   AryTypePara[234].Other.FixtureEnable := FALSE;
   AryTypePara[234].Other.Byte_1 := 16#00;
   AryTypePara[234].Other.Int_1 := 0;
   AryTypePara[234].Other."Char" := ' ';
   AryTypePara[234].Other.Word_1 := 16#0000;
   AryTypePara[234].Other.DInt_1 := 0;
   AryTypePara[234].Other.DWord_1 := 16#0000_0000;
   AryTypePara[234].Other.Real_1 := 0.0;
   AryTypePara[234].Other.S5Time := T#0MS;
   AryTypePara[234].Other."String" := '';
   AryTypePara[235].TypeName := '';
   AryTypePara[235].bit.Bit0 := FALSE;
   AryTypePara[235].bit.sp := 16#0000;
   AryTypePara[235].bit.Other.Bool_1 := FALSE;
   AryTypePara[235].bit.Other.Byte_2 := 16#00;
   AryTypePara[235].bit.Other.Int_1 := 0;
   AryTypePara[235].bit.Other."Char" := ' ';
   AryTypePara[235].Other.STxxxCCDProgNO := 0;
   AryTypePara[235].Other.FixtureEnable := FALSE;
   AryTypePara[235].Other.Byte_1 := 16#00;
   AryTypePara[235].Other.Int_1 := 0;
   AryTypePara[235].Other."Char" := ' ';
   AryTypePara[235].Other.Word_1 := 16#0000;
   AryTypePara[235].Other.DInt_1 := 0;
   AryTypePara[235].Other.DWord_1 := 16#0000_0000;
   AryTypePara[235].Other.Real_1 := 0.0;
   AryTypePara[235].Other.S5Time := T#0MS;
   AryTypePara[235].Other."String" := '';
   AryTypePara[236].TypeName := '';
   AryTypePara[236].bit.Bit0 := FALSE;
   AryTypePara[236].bit.sp := 16#0000;
   AryTypePara[236].bit.Other.Bool_1 := FALSE;
   AryTypePara[236].bit.Other.Byte_2 := 16#00;
   AryTypePara[236].bit.Other.Int_1 := 0;
   AryTypePara[236].bit.Other."Char" := ' ';
   AryTypePara[236].Other.STxxxCCDProgNO := 0;
   AryTypePara[236].Other.FixtureEnable := FALSE;
   AryTypePara[236].Other.Byte_1 := 16#00;
   AryTypePara[236].Other.Int_1 := 0;
   AryTypePara[236].Other."Char" := ' ';
   AryTypePara[236].Other.Word_1 := 16#0000;
   AryTypePara[236].Other.DInt_1 := 0;
   AryTypePara[236].Other.DWord_1 := 16#0000_0000;
   AryTypePara[236].Other.Real_1 := 0.0;
   AryTypePara[236].Other.S5Time := T#0MS;
   AryTypePara[236].Other."String" := '';
   AryTypePara[237].TypeName := '';
   AryTypePara[237].bit.Bit0 := FALSE;
   AryTypePara[237].bit.sp := 16#0000;
   AryTypePara[237].bit.Other.Bool_1 := FALSE;
   AryTypePara[237].bit.Other.Byte_2 := 16#00;
   AryTypePara[237].bit.Other.Int_1 := 0;
   AryTypePara[237].bit.Other."Char" := ' ';
   AryTypePara[237].Other.STxxxCCDProgNO := 0;
   AryTypePara[237].Other.FixtureEnable := FALSE;
   AryTypePara[237].Other.Byte_1 := 16#00;
   AryTypePara[237].Other.Int_1 := 0;
   AryTypePara[237].Other."Char" := ' ';
   AryTypePara[237].Other.Word_1 := 16#0000;
   AryTypePara[237].Other.DInt_1 := 0;
   AryTypePara[237].Other.DWord_1 := 16#0000_0000;
   AryTypePara[237].Other.Real_1 := 0.0;
   AryTypePara[237].Other.S5Time := T#0MS;
   AryTypePara[237].Other."String" := '';
   AryTypePara[238].TypeName := '';
   AryTypePara[238].bit.Bit0 := FALSE;
   AryTypePara[238].bit.sp := 16#0000;
   AryTypePara[238].bit.Other.Bool_1 := FALSE;
   AryTypePara[238].bit.Other.Byte_2 := 16#00;
   AryTypePara[238].bit.Other.Int_1 := 0;
   AryTypePara[238].bit.Other."Char" := ' ';
   AryTypePara[238].Other.STxxxCCDProgNO := 0;
   AryTypePara[238].Other.FixtureEnable := FALSE;
   AryTypePara[238].Other.Byte_1 := 16#00;
   AryTypePara[238].Other.Int_1 := 0;
   AryTypePara[238].Other."Char" := ' ';
   AryTypePara[238].Other.Word_1 := 16#0000;
   AryTypePara[238].Other.DInt_1 := 0;
   AryTypePara[238].Other.DWord_1 := 16#0000_0000;
   AryTypePara[238].Other.Real_1 := 0.0;
   AryTypePara[238].Other.S5Time := T#0MS;
   AryTypePara[238].Other."String" := '';
   AryTypePara[239].TypeName := '';
   AryTypePara[239].bit.Bit0 := FALSE;
   AryTypePara[239].bit.sp := 16#0000;
   AryTypePara[239].bit.Other.Bool_1 := FALSE;
   AryTypePara[239].bit.Other.Byte_2 := 16#00;
   AryTypePara[239].bit.Other.Int_1 := 0;
   AryTypePara[239].bit.Other."Char" := ' ';
   AryTypePara[239].Other.STxxxCCDProgNO := 0;
   AryTypePara[239].Other.FixtureEnable := FALSE;
   AryTypePara[239].Other.Byte_1 := 16#00;
   AryTypePara[239].Other.Int_1 := 0;
   AryTypePara[239].Other."Char" := ' ';
   AryTypePara[239].Other.Word_1 := 16#0000;
   AryTypePara[239].Other.DInt_1 := 0;
   AryTypePara[239].Other.DWord_1 := 16#0000_0000;
   AryTypePara[239].Other.Real_1 := 0.0;
   AryTypePara[239].Other.S5Time := T#0MS;
   AryTypePara[239].Other."String" := '';
   AryTypePara[240].TypeName := '';
   AryTypePara[240].bit.Bit0 := FALSE;
   AryTypePara[240].bit.sp := 16#0000;
   AryTypePara[240].bit.Other.Bool_1 := FALSE;
   AryTypePara[240].bit.Other.Byte_2 := 16#00;
   AryTypePara[240].bit.Other.Int_1 := 0;
   AryTypePara[240].bit.Other."Char" := ' ';
   AryTypePara[240].Other.STxxxCCDProgNO := 0;
   AryTypePara[240].Other.FixtureEnable := FALSE;
   AryTypePara[240].Other.Byte_1 := 16#00;
   AryTypePara[240].Other.Int_1 := 0;
   AryTypePara[240].Other."Char" := ' ';
   AryTypePara[240].Other.Word_1 := 16#0000;
   AryTypePara[240].Other.DInt_1 := 0;
   AryTypePara[240].Other.DWord_1 := 16#0000_0000;
   AryTypePara[240].Other.Real_1 := 0.0;
   AryTypePara[240].Other.S5Time := T#0MS;
   AryTypePara[240].Other."String" := '';
   AryTypePara[241].TypeName := '';
   AryTypePara[241].bit.Bit0 := FALSE;
   AryTypePara[241].bit.sp := 16#0000;
   AryTypePara[241].bit.Other.Bool_1 := FALSE;
   AryTypePara[241].bit.Other.Byte_2 := 16#00;
   AryTypePara[241].bit.Other.Int_1 := 0;
   AryTypePara[241].bit.Other."Char" := ' ';
   AryTypePara[241].Other.STxxxCCDProgNO := 0;
   AryTypePara[241].Other.FixtureEnable := FALSE;
   AryTypePara[241].Other.Byte_1 := 16#00;
   AryTypePara[241].Other.Int_1 := 0;
   AryTypePara[241].Other."Char" := ' ';
   AryTypePara[241].Other.Word_1 := 16#0000;
   AryTypePara[241].Other.DInt_1 := 0;
   AryTypePara[241].Other.DWord_1 := 16#0000_0000;
   AryTypePara[241].Other.Real_1 := 0.0;
   AryTypePara[241].Other.S5Time := T#0MS;
   AryTypePara[241].Other."String" := '';
   AryTypePara[242].TypeName := '';
   AryTypePara[242].bit.Bit0 := FALSE;
   AryTypePara[242].bit.sp := 16#0000;
   AryTypePara[242].bit.Other.Bool_1 := FALSE;
   AryTypePara[242].bit.Other.Byte_2 := 16#00;
   AryTypePara[242].bit.Other.Int_1 := 0;
   AryTypePara[242].bit.Other."Char" := ' ';
   AryTypePara[242].Other.STxxxCCDProgNO := 0;
   AryTypePara[242].Other.FixtureEnable := FALSE;
   AryTypePara[242].Other.Byte_1 := 16#00;
   AryTypePara[242].Other.Int_1 := 0;
   AryTypePara[242].Other."Char" := ' ';
   AryTypePara[242].Other.Word_1 := 16#0000;
   AryTypePara[242].Other.DInt_1 := 0;
   AryTypePara[242].Other.DWord_1 := 16#0000_0000;
   AryTypePara[242].Other.Real_1 := 0.0;
   AryTypePara[242].Other.S5Time := T#0MS;
   AryTypePara[242].Other."String" := '';
   AryTypePara[243].TypeName := '';
   AryTypePara[243].bit.Bit0 := FALSE;
   AryTypePara[243].bit.sp := 16#0000;
   AryTypePara[243].bit.Other.Bool_1 := FALSE;
   AryTypePara[243].bit.Other.Byte_2 := 16#00;
   AryTypePara[243].bit.Other.Int_1 := 0;
   AryTypePara[243].bit.Other."Char" := ' ';
   AryTypePara[243].Other.STxxxCCDProgNO := 0;
   AryTypePara[243].Other.FixtureEnable := FALSE;
   AryTypePara[243].Other.Byte_1 := 16#00;
   AryTypePara[243].Other.Int_1 := 0;
   AryTypePara[243].Other."Char" := ' ';
   AryTypePara[243].Other.Word_1 := 16#0000;
   AryTypePara[243].Other.DInt_1 := 0;
   AryTypePara[243].Other.DWord_1 := 16#0000_0000;
   AryTypePara[243].Other.Real_1 := 0.0;
   AryTypePara[243].Other.S5Time := T#0MS;
   AryTypePara[243].Other."String" := '';
   AryTypePara[244].TypeName := '';
   AryTypePara[244].bit.Bit0 := FALSE;
   AryTypePara[244].bit.sp := 16#0000;
   AryTypePara[244].bit.Other.Bool_1 := FALSE;
   AryTypePara[244].bit.Other.Byte_2 := 16#00;
   AryTypePara[244].bit.Other.Int_1 := 0;
   AryTypePara[244].bit.Other."Char" := ' ';
   AryTypePara[244].Other.STxxxCCDProgNO := 0;
   AryTypePara[244].Other.FixtureEnable := FALSE;
   AryTypePara[244].Other.Byte_1 := 16#00;
   AryTypePara[244].Other.Int_1 := 0;
   AryTypePara[244].Other."Char" := ' ';
   AryTypePara[244].Other.Word_1 := 16#0000;
   AryTypePara[244].Other.DInt_1 := 0;
   AryTypePara[244].Other.DWord_1 := 16#0000_0000;
   AryTypePara[244].Other.Real_1 := 0.0;
   AryTypePara[244].Other.S5Time := T#0MS;
   AryTypePara[244].Other."String" := '';
   AryTypePara[245].TypeName := '';
   AryTypePara[245].bit.Bit0 := FALSE;
   AryTypePara[245].bit.sp := 16#0000;
   AryTypePara[245].bit.Other.Bool_1 := FALSE;
   AryTypePara[245].bit.Other.Byte_2 := 16#00;
   AryTypePara[245].bit.Other.Int_1 := 0;
   AryTypePara[245].bit.Other."Char" := ' ';
   AryTypePara[245].Other.STxxxCCDProgNO := 0;
   AryTypePara[245].Other.FixtureEnable := FALSE;
   AryTypePara[245].Other.Byte_1 := 16#00;
   AryTypePara[245].Other.Int_1 := 0;
   AryTypePara[245].Other."Char" := ' ';
   AryTypePara[245].Other.Word_1 := 16#0000;
   AryTypePara[245].Other.DInt_1 := 0;
   AryTypePara[245].Other.DWord_1 := 16#0000_0000;
   AryTypePara[245].Other.Real_1 := 0.0;
   AryTypePara[245].Other.S5Time := T#0MS;
   AryTypePara[245].Other."String" := '';
   AryTypePara[246].TypeName := '';
   AryTypePara[246].bit.Bit0 := FALSE;
   AryTypePara[246].bit.sp := 16#0000;
   AryTypePara[246].bit.Other.Bool_1 := FALSE;
   AryTypePara[246].bit.Other.Byte_2 := 16#00;
   AryTypePara[246].bit.Other.Int_1 := 0;
   AryTypePara[246].bit.Other."Char" := ' ';
   AryTypePara[246].Other.STxxxCCDProgNO := 0;
   AryTypePara[246].Other.FixtureEnable := FALSE;
   AryTypePara[246].Other.Byte_1 := 16#00;
   AryTypePara[246].Other.Int_1 := 0;
   AryTypePara[246].Other."Char" := ' ';
   AryTypePara[246].Other.Word_1 := 16#0000;
   AryTypePara[246].Other.DInt_1 := 0;
   AryTypePara[246].Other.DWord_1 := 16#0000_0000;
   AryTypePara[246].Other.Real_1 := 0.0;
   AryTypePara[246].Other.S5Time := T#0MS;
   AryTypePara[246].Other."String" := '';
   AryTypePara[247].TypeName := '';
   AryTypePara[247].bit.Bit0 := FALSE;
   AryTypePara[247].bit.sp := 16#0000;
   AryTypePara[247].bit.Other.Bool_1 := FALSE;
   AryTypePara[247].bit.Other.Byte_2 := 16#00;
   AryTypePara[247].bit.Other.Int_1 := 0;
   AryTypePara[247].bit.Other."Char" := ' ';
   AryTypePara[247].Other.STxxxCCDProgNO := 0;
   AryTypePara[247].Other.FixtureEnable := FALSE;
   AryTypePara[247].Other.Byte_1 := 16#00;
   AryTypePara[247].Other.Int_1 := 0;
   AryTypePara[247].Other."Char" := ' ';
   AryTypePara[247].Other.Word_1 := 16#0000;
   AryTypePara[247].Other.DInt_1 := 0;
   AryTypePara[247].Other.DWord_1 := 16#0000_0000;
   AryTypePara[247].Other.Real_1 := 0.0;
   AryTypePara[247].Other.S5Time := T#0MS;
   AryTypePara[247].Other."String" := '';
   AryTypePara[248].TypeName := '';
   AryTypePara[248].bit.Bit0 := FALSE;
   AryTypePara[248].bit.sp := 16#0000;
   AryTypePara[248].bit.Other.Bool_1 := FALSE;
   AryTypePara[248].bit.Other.Byte_2 := 16#00;
   AryTypePara[248].bit.Other.Int_1 := 0;
   AryTypePara[248].bit.Other."Char" := ' ';
   AryTypePara[248].Other.STxxxCCDProgNO := 0;
   AryTypePara[248].Other.FixtureEnable := FALSE;
   AryTypePara[248].Other.Byte_1 := 16#00;
   AryTypePara[248].Other.Int_1 := 0;
   AryTypePara[248].Other."Char" := ' ';
   AryTypePara[248].Other.Word_1 := 16#0000;
   AryTypePara[248].Other.DInt_1 := 0;
   AryTypePara[248].Other.DWord_1 := 16#0000_0000;
   AryTypePara[248].Other.Real_1 := 0.0;
   AryTypePara[248].Other.S5Time := T#0MS;
   AryTypePara[248].Other."String" := '';
   AryTypePara[249].TypeName := '';
   AryTypePara[249].bit.Bit0 := FALSE;
   AryTypePara[249].bit.sp := 16#0000;
   AryTypePara[249].bit.Other.Bool_1 := FALSE;
   AryTypePara[249].bit.Other.Byte_2 := 16#00;
   AryTypePara[249].bit.Other.Int_1 := 0;
   AryTypePara[249].bit.Other."Char" := ' ';
   AryTypePara[249].Other.STxxxCCDProgNO := 0;
   AryTypePara[249].Other.FixtureEnable := FALSE;
   AryTypePara[249].Other.Byte_1 := 16#00;
   AryTypePara[249].Other.Int_1 := 0;
   AryTypePara[249].Other."Char" := ' ';
   AryTypePara[249].Other.Word_1 := 16#0000;
   AryTypePara[249].Other.DInt_1 := 0;
   AryTypePara[249].Other.DWord_1 := 16#0000_0000;
   AryTypePara[249].Other.Real_1 := 0.0;
   AryTypePara[249].Other.S5Time := T#0MS;
   AryTypePara[249].Other."String" := '';
   AryTypePara[250].TypeName := '';
   AryTypePara[250].bit.Bit0 := FALSE;
   AryTypePara[250].bit.sp := 16#0000;
   AryTypePara[250].bit.Other.Bool_1 := FALSE;
   AryTypePara[250].bit.Other.Byte_2 := 16#00;
   AryTypePara[250].bit.Other.Int_1 := 0;
   AryTypePara[250].bit.Other."Char" := ' ';
   AryTypePara[250].Other.STxxxCCDProgNO := 0;
   AryTypePara[250].Other.FixtureEnable := FALSE;
   AryTypePara[250].Other.Byte_1 := 16#00;
   AryTypePara[250].Other.Int_1 := 0;
   AryTypePara[250].Other."Char" := ' ';
   AryTypePara[250].Other.Word_1 := 16#0000;
   AryTypePara[250].Other.DInt_1 := 0;
   AryTypePara[250].Other.DWord_1 := 16#0000_0000;
   AryTypePara[250].Other.Real_1 := 0.0;
   AryTypePara[250].Other.S5Time := T#0MS;
   AryTypePara[250].Other."String" := '';
   AryTypePara[251].TypeName := '';
   AryTypePara[251].bit.Bit0 := FALSE;
   AryTypePara[251].bit.sp := 16#0000;
   AryTypePara[251].bit.Other.Bool_1 := FALSE;
   AryTypePara[251].bit.Other.Byte_2 := 16#00;
   AryTypePara[251].bit.Other.Int_1 := 0;
   AryTypePara[251].bit.Other."Char" := ' ';
   AryTypePara[251].Other.STxxxCCDProgNO := 0;
   AryTypePara[251].Other.FixtureEnable := FALSE;
   AryTypePara[251].Other.Byte_1 := 16#00;
   AryTypePara[251].Other.Int_1 := 0;
   AryTypePara[251].Other."Char" := ' ';
   AryTypePara[251].Other.Word_1 := 16#0000;
   AryTypePara[251].Other.DInt_1 := 0;
   AryTypePara[251].Other.DWord_1 := 16#0000_0000;
   AryTypePara[251].Other.Real_1 := 0.0;
   AryTypePara[251].Other.S5Time := T#0MS;
   AryTypePara[251].Other."String" := '';
   AryTypePara[252].TypeName := '';
   AryTypePara[252].bit.Bit0 := FALSE;
   AryTypePara[252].bit.sp := 16#0000;
   AryTypePara[252].bit.Other.Bool_1 := FALSE;
   AryTypePara[252].bit.Other.Byte_2 := 16#00;
   AryTypePara[252].bit.Other.Int_1 := 0;
   AryTypePara[252].bit.Other."Char" := ' ';
   AryTypePara[252].Other.STxxxCCDProgNO := 0;
   AryTypePara[252].Other.FixtureEnable := FALSE;
   AryTypePara[252].Other.Byte_1 := 16#00;
   AryTypePara[252].Other.Int_1 := 0;
   AryTypePara[252].Other."Char" := ' ';
   AryTypePara[252].Other.Word_1 := 16#0000;
   AryTypePara[252].Other.DInt_1 := 0;
   AryTypePara[252].Other.DWord_1 := 16#0000_0000;
   AryTypePara[252].Other.Real_1 := 0.0;
   AryTypePara[252].Other.S5Time := T#0MS;
   AryTypePara[252].Other."String" := '';
   AryTypePara[253].TypeName := '';
   AryTypePara[253].bit.Bit0 := FALSE;
   AryTypePara[253].bit.sp := 16#0000;
   AryTypePara[253].bit.Other.Bool_1 := FALSE;
   AryTypePara[253].bit.Other.Byte_2 := 16#00;
   AryTypePara[253].bit.Other.Int_1 := 0;
   AryTypePara[253].bit.Other."Char" := ' ';
   AryTypePara[253].Other.STxxxCCDProgNO := 0;
   AryTypePara[253].Other.FixtureEnable := FALSE;
   AryTypePara[253].Other.Byte_1 := 16#00;
   AryTypePara[253].Other.Int_1 := 0;
   AryTypePara[253].Other."Char" := ' ';
   AryTypePara[253].Other.Word_1 := 16#0000;
   AryTypePara[253].Other.DInt_1 := 0;
   AryTypePara[253].Other.DWord_1 := 16#0000_0000;
   AryTypePara[253].Other.Real_1 := 0.0;
   AryTypePara[253].Other.S5Time := T#0MS;
   AryTypePara[253].Other."String" := '';
   AryTypePara[254].TypeName := '';
   AryTypePara[254].bit.Bit0 := FALSE;
   AryTypePara[254].bit.sp := 16#0000;
   AryTypePara[254].bit.Other.Bool_1 := FALSE;
   AryTypePara[254].bit.Other.Byte_2 := 16#00;
   AryTypePara[254].bit.Other.Int_1 := 0;
   AryTypePara[254].bit.Other."Char" := ' ';
   AryTypePara[254].Other.STxxxCCDProgNO := 0;
   AryTypePara[254].Other.FixtureEnable := FALSE;
   AryTypePara[254].Other.Byte_1 := 16#00;
   AryTypePara[254].Other.Int_1 := 0;
   AryTypePara[254].Other."Char" := ' ';
   AryTypePara[254].Other.Word_1 := 16#0000;
   AryTypePara[254].Other.DInt_1 := 0;
   AryTypePara[254].Other.DWord_1 := 16#0000_0000;
   AryTypePara[254].Other.Real_1 := 0.0;
   AryTypePara[254].Other.S5Time := T#0MS;
   AryTypePara[254].Other."String" := '';
   AryTypePara[255].TypeName := '';
   AryTypePara[255].bit.Bit0 := FALSE;
   AryTypePara[255].bit.sp := 16#0000;
   AryTypePara[255].bit.Other.Bool_1 := FALSE;
   AryTypePara[255].bit.Other.Byte_2 := 16#00;
   AryTypePara[255].bit.Other.Int_1 := 0;
   AryTypePara[255].bit.Other."Char" := ' ';
   AryTypePara[255].Other.STxxxCCDProgNO := 0;
   AryTypePara[255].Other.FixtureEnable := FALSE;
   AryTypePara[255].Other.Byte_1 := 16#00;
   AryTypePara[255].Other.Int_1 := 0;
   AryTypePara[255].Other."Char" := ' ';
   AryTypePara[255].Other.Word_1 := 16#0000;
   AryTypePara[255].Other.DInt_1 := 0;
   AryTypePara[255].Other.DWord_1 := 16#0000_0000;
   AryTypePara[255].Other.Real_1 := 0.0;
   AryTypePara[255].Other.S5Time := T#0MS;
   AryTypePara[255].Other."String" := '';
   AryTypePara[256].TypeName := '';
   AryTypePara[256].bit.Bit0 := FALSE;
   AryTypePara[256].bit.sp := 16#0000;
   AryTypePara[256].bit.Other.Bool_1 := FALSE;
   AryTypePara[256].bit.Other.Byte_2 := 16#00;
   AryTypePara[256].bit.Other.Int_1 := 0;
   AryTypePara[256].bit.Other."Char" := ' ';
   AryTypePara[256].Other.STxxxCCDProgNO := 0;
   AryTypePara[256].Other.FixtureEnable := FALSE;
   AryTypePara[256].Other.Byte_1 := 16#00;
   AryTypePara[256].Other.Int_1 := 0;
   AryTypePara[256].Other."Char" := ' ';
   AryTypePara[256].Other.Word_1 := 16#0000;
   AryTypePara[256].Other.DInt_1 := 0;
   AryTypePara[256].Other.DWord_1 := 16#0000_0000;
   AryTypePara[256].Other.Real_1 := 0.0;
   AryTypePara[256].Other.S5Time := T#0MS;
   AryTypePara[256].Other."String" := '';
   AryTypePara[257].TypeName := '';
   AryTypePara[257].bit.Bit0 := FALSE;
   AryTypePara[257].bit.sp := 16#0000;
   AryTypePara[257].bit.Other.Bool_1 := FALSE;
   AryTypePara[257].bit.Other.Byte_2 := 16#00;
   AryTypePara[257].bit.Other.Int_1 := 0;
   AryTypePara[257].bit.Other."Char" := ' ';
   AryTypePara[257].Other.STxxxCCDProgNO := 0;
   AryTypePara[257].Other.FixtureEnable := FALSE;
   AryTypePara[257].Other.Byte_1 := 16#00;
   AryTypePara[257].Other.Int_1 := 0;
   AryTypePara[257].Other."Char" := ' ';
   AryTypePara[257].Other.Word_1 := 16#0000;
   AryTypePara[257].Other.DInt_1 := 0;
   AryTypePara[257].Other.DWord_1 := 16#0000_0000;
   AryTypePara[257].Other.Real_1 := 0.0;
   AryTypePara[257].Other.S5Time := T#0MS;
   AryTypePara[257].Other."String" := '';
   AryTypePara[258].TypeName := '';
   AryTypePara[258].bit.Bit0 := FALSE;
   AryTypePara[258].bit.sp := 16#0000;
   AryTypePara[258].bit.Other.Bool_1 := FALSE;
   AryTypePara[258].bit.Other.Byte_2 := 16#00;
   AryTypePara[258].bit.Other.Int_1 := 0;
   AryTypePara[258].bit.Other."Char" := ' ';
   AryTypePara[258].Other.STxxxCCDProgNO := 0;
   AryTypePara[258].Other.FixtureEnable := FALSE;
   AryTypePara[258].Other.Byte_1 := 16#00;
   AryTypePara[258].Other.Int_1 := 0;
   AryTypePara[258].Other."Char" := ' ';
   AryTypePara[258].Other.Word_1 := 16#0000;
   AryTypePara[258].Other.DInt_1 := 0;
   AryTypePara[258].Other.DWord_1 := 16#0000_0000;
   AryTypePara[258].Other.Real_1 := 0.0;
   AryTypePara[258].Other.S5Time := T#0MS;
   AryTypePara[258].Other."String" := '';
   AryTypePara[259].TypeName := '';
   AryTypePara[259].bit.Bit0 := FALSE;
   AryTypePara[259].bit.sp := 16#0000;
   AryTypePara[259].bit.Other.Bool_1 := FALSE;
   AryTypePara[259].bit.Other.Byte_2 := 16#00;
   AryTypePara[259].bit.Other.Int_1 := 0;
   AryTypePara[259].bit.Other."Char" := ' ';
   AryTypePara[259].Other.STxxxCCDProgNO := 0;
   AryTypePara[259].Other.FixtureEnable := FALSE;
   AryTypePara[259].Other.Byte_1 := 16#00;
   AryTypePara[259].Other.Int_1 := 0;
   AryTypePara[259].Other."Char" := ' ';
   AryTypePara[259].Other.Word_1 := 16#0000;
   AryTypePara[259].Other.DInt_1 := 0;
   AryTypePara[259].Other.DWord_1 := 16#0000_0000;
   AryTypePara[259].Other.Real_1 := 0.0;
   AryTypePara[259].Other.S5Time := T#0MS;
   AryTypePara[259].Other."String" := '';
   AryTypePara[260].TypeName := '';
   AryTypePara[260].bit.Bit0 := FALSE;
   AryTypePara[260].bit.sp := 16#0000;
   AryTypePara[260].bit.Other.Bool_1 := FALSE;
   AryTypePara[260].bit.Other.Byte_2 := 16#00;
   AryTypePara[260].bit.Other.Int_1 := 0;
   AryTypePara[260].bit.Other."Char" := ' ';
   AryTypePara[260].Other.STxxxCCDProgNO := 0;
   AryTypePara[260].Other.FixtureEnable := FALSE;
   AryTypePara[260].Other.Byte_1 := 16#00;
   AryTypePara[260].Other.Int_1 := 0;
   AryTypePara[260].Other."Char" := ' ';
   AryTypePara[260].Other.Word_1 := 16#0000;
   AryTypePara[260].Other.DInt_1 := 0;
   AryTypePara[260].Other.DWord_1 := 16#0000_0000;
   AryTypePara[260].Other.Real_1 := 0.0;
   AryTypePara[260].Other.S5Time := T#0MS;
   AryTypePara[260].Other."String" := '';
   AryTypePara[261].TypeName := '';
   AryTypePara[261].bit.Bit0 := FALSE;
   AryTypePara[261].bit.sp := 16#0000;
   AryTypePara[261].bit.Other.Bool_1 := FALSE;
   AryTypePara[261].bit.Other.Byte_2 := 16#00;
   AryTypePara[261].bit.Other.Int_1 := 0;
   AryTypePara[261].bit.Other."Char" := ' ';
   AryTypePara[261].Other.STxxxCCDProgNO := 0;
   AryTypePara[261].Other.FixtureEnable := FALSE;
   AryTypePara[261].Other.Byte_1 := 16#00;
   AryTypePara[261].Other.Int_1 := 0;
   AryTypePara[261].Other."Char" := ' ';
   AryTypePara[261].Other.Word_1 := 16#0000;
   AryTypePara[261].Other.DInt_1 := 0;
   AryTypePara[261].Other.DWord_1 := 16#0000_0000;
   AryTypePara[261].Other.Real_1 := 0.0;
   AryTypePara[261].Other.S5Time := T#0MS;
   AryTypePara[261].Other."String" := '';
   AryTypePara[262].TypeName := '';
   AryTypePara[262].bit.Bit0 := FALSE;
   AryTypePara[262].bit.sp := 16#0000;
   AryTypePara[262].bit.Other.Bool_1 := FALSE;
   AryTypePara[262].bit.Other.Byte_2 := 16#00;
   AryTypePara[262].bit.Other.Int_1 := 0;
   AryTypePara[262].bit.Other."Char" := ' ';
   AryTypePara[262].Other.STxxxCCDProgNO := 0;
   AryTypePara[262].Other.FixtureEnable := FALSE;
   AryTypePara[262].Other.Byte_1 := 16#00;
   AryTypePara[262].Other.Int_1 := 0;
   AryTypePara[262].Other."Char" := ' ';
   AryTypePara[262].Other.Word_1 := 16#0000;
   AryTypePara[262].Other.DInt_1 := 0;
   AryTypePara[262].Other.DWord_1 := 16#0000_0000;
   AryTypePara[262].Other.Real_1 := 0.0;
   AryTypePara[262].Other.S5Time := T#0MS;
   AryTypePara[262].Other."String" := '';
   AryTypePara[263].TypeName := '';
   AryTypePara[263].bit.Bit0 := FALSE;
   AryTypePara[263].bit.sp := 16#0000;
   AryTypePara[263].bit.Other.Bool_1 := FALSE;
   AryTypePara[263].bit.Other.Byte_2 := 16#00;
   AryTypePara[263].bit.Other.Int_1 := 0;
   AryTypePara[263].bit.Other."Char" := ' ';
   AryTypePara[263].Other.STxxxCCDProgNO := 0;
   AryTypePara[263].Other.FixtureEnable := FALSE;
   AryTypePara[263].Other.Byte_1 := 16#00;
   AryTypePara[263].Other.Int_1 := 0;
   AryTypePara[263].Other."Char" := ' ';
   AryTypePara[263].Other.Word_1 := 16#0000;
   AryTypePara[263].Other.DInt_1 := 0;
   AryTypePara[263].Other.DWord_1 := 16#0000_0000;
   AryTypePara[263].Other.Real_1 := 0.0;
   AryTypePara[263].Other.S5Time := T#0MS;
   AryTypePara[263].Other."String" := '';
   AryTypePara[264].TypeName := '';
   AryTypePara[264].bit.Bit0 := FALSE;
   AryTypePara[264].bit.sp := 16#0000;
   AryTypePara[264].bit.Other.Bool_1 := FALSE;
   AryTypePara[264].bit.Other.Byte_2 := 16#00;
   AryTypePara[264].bit.Other.Int_1 := 0;
   AryTypePara[264].bit.Other."Char" := ' ';
   AryTypePara[264].Other.STxxxCCDProgNO := 0;
   AryTypePara[264].Other.FixtureEnable := FALSE;
   AryTypePara[264].Other.Byte_1 := 16#00;
   AryTypePara[264].Other.Int_1 := 0;
   AryTypePara[264].Other."Char" := ' ';
   AryTypePara[264].Other.Word_1 := 16#0000;
   AryTypePara[264].Other.DInt_1 := 0;
   AryTypePara[264].Other.DWord_1 := 16#0000_0000;
   AryTypePara[264].Other.Real_1 := 0.0;
   AryTypePara[264].Other.S5Time := T#0MS;
   AryTypePara[264].Other."String" := '';
   AryTypePara[265].TypeName := '';
   AryTypePara[265].bit.Bit0 := FALSE;
   AryTypePara[265].bit.sp := 16#0000;
   AryTypePara[265].bit.Other.Bool_1 := FALSE;
   AryTypePara[265].bit.Other.Byte_2 := 16#00;
   AryTypePara[265].bit.Other.Int_1 := 0;
   AryTypePara[265].bit.Other."Char" := ' ';
   AryTypePara[265].Other.STxxxCCDProgNO := 0;
   AryTypePara[265].Other.FixtureEnable := FALSE;
   AryTypePara[265].Other.Byte_1 := 16#00;
   AryTypePara[265].Other.Int_1 := 0;
   AryTypePara[265].Other."Char" := ' ';
   AryTypePara[265].Other.Word_1 := 16#0000;
   AryTypePara[265].Other.DInt_1 := 0;
   AryTypePara[265].Other.DWord_1 := 16#0000_0000;
   AryTypePara[265].Other.Real_1 := 0.0;
   AryTypePara[265].Other.S5Time := T#0MS;
   AryTypePara[265].Other."String" := '';
   AryTypePara[266].TypeName := '';
   AryTypePara[266].bit.Bit0 := FALSE;
   AryTypePara[266].bit.sp := 16#0000;
   AryTypePara[266].bit.Other.Bool_1 := FALSE;
   AryTypePara[266].bit.Other.Byte_2 := 16#00;
   AryTypePara[266].bit.Other.Int_1 := 0;
   AryTypePara[266].bit.Other."Char" := ' ';
   AryTypePara[266].Other.STxxxCCDProgNO := 0;
   AryTypePara[266].Other.FixtureEnable := FALSE;
   AryTypePara[266].Other.Byte_1 := 16#00;
   AryTypePara[266].Other.Int_1 := 0;
   AryTypePara[266].Other."Char" := ' ';
   AryTypePara[266].Other.Word_1 := 16#0000;
   AryTypePara[266].Other.DInt_1 := 0;
   AryTypePara[266].Other.DWord_1 := 16#0000_0000;
   AryTypePara[266].Other.Real_1 := 0.0;
   AryTypePara[266].Other.S5Time := T#0MS;
   AryTypePara[266].Other."String" := '';
   AryTypePara[267].TypeName := '';
   AryTypePara[267].bit.Bit0 := FALSE;
   AryTypePara[267].bit.sp := 16#0000;
   AryTypePara[267].bit.Other.Bool_1 := FALSE;
   AryTypePara[267].bit.Other.Byte_2 := 16#00;
   AryTypePara[267].bit.Other.Int_1 := 0;
   AryTypePara[267].bit.Other."Char" := ' ';
   AryTypePara[267].Other.STxxxCCDProgNO := 0;
   AryTypePara[267].Other.FixtureEnable := FALSE;
   AryTypePara[267].Other.Byte_1 := 16#00;
   AryTypePara[267].Other.Int_1 := 0;
   AryTypePara[267].Other."Char" := ' ';
   AryTypePara[267].Other.Word_1 := 16#0000;
   AryTypePara[267].Other.DInt_1 := 0;
   AryTypePara[267].Other.DWord_1 := 16#0000_0000;
   AryTypePara[267].Other.Real_1 := 0.0;
   AryTypePara[267].Other.S5Time := T#0MS;
   AryTypePara[267].Other."String" := '';
   AryTypePara[268].TypeName := '';
   AryTypePara[268].bit.Bit0 := FALSE;
   AryTypePara[268].bit.sp := 16#0000;
   AryTypePara[268].bit.Other.Bool_1 := FALSE;
   AryTypePara[268].bit.Other.Byte_2 := 16#00;
   AryTypePara[268].bit.Other.Int_1 := 0;
   AryTypePara[268].bit.Other."Char" := ' ';
   AryTypePara[268].Other.STxxxCCDProgNO := 0;
   AryTypePara[268].Other.FixtureEnable := FALSE;
   AryTypePara[268].Other.Byte_1 := 16#00;
   AryTypePara[268].Other.Int_1 := 0;
   AryTypePara[268].Other."Char" := ' ';
   AryTypePara[268].Other.Word_1 := 16#0000;
   AryTypePara[268].Other.DInt_1 := 0;
   AryTypePara[268].Other.DWord_1 := 16#0000_0000;
   AryTypePara[268].Other.Real_1 := 0.0;
   AryTypePara[268].Other.S5Time := T#0MS;
   AryTypePara[268].Other."String" := '';
   AryTypePara[269].TypeName := '';
   AryTypePara[269].bit.Bit0 := FALSE;
   AryTypePara[269].bit.sp := 16#0000;
   AryTypePara[269].bit.Other.Bool_1 := FALSE;
   AryTypePara[269].bit.Other.Byte_2 := 16#00;
   AryTypePara[269].bit.Other.Int_1 := 0;
   AryTypePara[269].bit.Other."Char" := ' ';
   AryTypePara[269].Other.STxxxCCDProgNO := 0;
   AryTypePara[269].Other.FixtureEnable := FALSE;
   AryTypePara[269].Other.Byte_1 := 16#00;
   AryTypePara[269].Other.Int_1 := 0;
   AryTypePara[269].Other."Char" := ' ';
   AryTypePara[269].Other.Word_1 := 16#0000;
   AryTypePara[269].Other.DInt_1 := 0;
   AryTypePara[269].Other.DWord_1 := 16#0000_0000;
   AryTypePara[269].Other.Real_1 := 0.0;
   AryTypePara[269].Other.S5Time := T#0MS;
   AryTypePara[269].Other."String" := '';
   AryTypePara[270].TypeName := '';
   AryTypePara[270].bit.Bit0 := FALSE;
   AryTypePara[270].bit.sp := 16#0000;
   AryTypePara[270].bit.Other.Bool_1 := FALSE;
   AryTypePara[270].bit.Other.Byte_2 := 16#00;
   AryTypePara[270].bit.Other.Int_1 := 0;
   AryTypePara[270].bit.Other."Char" := ' ';
   AryTypePara[270].Other.STxxxCCDProgNO := 0;
   AryTypePara[270].Other.FixtureEnable := FALSE;
   AryTypePara[270].Other.Byte_1 := 16#00;
   AryTypePara[270].Other.Int_1 := 0;
   AryTypePara[270].Other."Char" := ' ';
   AryTypePara[270].Other.Word_1 := 16#0000;
   AryTypePara[270].Other.DInt_1 := 0;
   AryTypePara[270].Other.DWord_1 := 16#0000_0000;
   AryTypePara[270].Other.Real_1 := 0.0;
   AryTypePara[270].Other.S5Time := T#0MS;
   AryTypePara[270].Other."String" := '';
   AryTypePara[271].TypeName := '';
   AryTypePara[271].bit.Bit0 := FALSE;
   AryTypePara[271].bit.sp := 16#0000;
   AryTypePara[271].bit.Other.Bool_1 := FALSE;
   AryTypePara[271].bit.Other.Byte_2 := 16#00;
   AryTypePara[271].bit.Other.Int_1 := 0;
   AryTypePara[271].bit.Other."Char" := ' ';
   AryTypePara[271].Other.STxxxCCDProgNO := 0;
   AryTypePara[271].Other.FixtureEnable := FALSE;
   AryTypePara[271].Other.Byte_1 := 16#00;
   AryTypePara[271].Other.Int_1 := 0;
   AryTypePara[271].Other."Char" := ' ';
   AryTypePara[271].Other.Word_1 := 16#0000;
   AryTypePara[271].Other.DInt_1 := 0;
   AryTypePara[271].Other.DWord_1 := 16#0000_0000;
   AryTypePara[271].Other.Real_1 := 0.0;
   AryTypePara[271].Other.S5Time := T#0MS;
   AryTypePara[271].Other."String" := '';
   AryTypePara[272].TypeName := '';
   AryTypePara[272].bit.Bit0 := FALSE;
   AryTypePara[272].bit.sp := 16#0000;
   AryTypePara[272].bit.Other.Bool_1 := FALSE;
   AryTypePara[272].bit.Other.Byte_2 := 16#00;
   AryTypePara[272].bit.Other.Int_1 := 0;
   AryTypePara[272].bit.Other."Char" := ' ';
   AryTypePara[272].Other.STxxxCCDProgNO := 0;
   AryTypePara[272].Other.FixtureEnable := FALSE;
   AryTypePara[272].Other.Byte_1 := 16#00;
   AryTypePara[272].Other.Int_1 := 0;
   AryTypePara[272].Other."Char" := ' ';
   AryTypePara[272].Other.Word_1 := 16#0000;
   AryTypePara[272].Other.DInt_1 := 0;
   AryTypePara[272].Other.DWord_1 := 16#0000_0000;
   AryTypePara[272].Other.Real_1 := 0.0;
   AryTypePara[272].Other.S5Time := T#0MS;
   AryTypePara[272].Other."String" := '';
   AryTypePara[273].TypeName := '';
   AryTypePara[273].bit.Bit0 := FALSE;
   AryTypePara[273].bit.sp := 16#0000;
   AryTypePara[273].bit.Other.Bool_1 := FALSE;
   AryTypePara[273].bit.Other.Byte_2 := 16#00;
   AryTypePara[273].bit.Other.Int_1 := 0;
   AryTypePara[273].bit.Other."Char" := ' ';
   AryTypePara[273].Other.STxxxCCDProgNO := 0;
   AryTypePara[273].Other.FixtureEnable := FALSE;
   AryTypePara[273].Other.Byte_1 := 16#00;
   AryTypePara[273].Other.Int_1 := 0;
   AryTypePara[273].Other."Char" := ' ';
   AryTypePara[273].Other.Word_1 := 16#0000;
   AryTypePara[273].Other.DInt_1 := 0;
   AryTypePara[273].Other.DWord_1 := 16#0000_0000;
   AryTypePara[273].Other.Real_1 := 0.0;
   AryTypePara[273].Other.S5Time := T#0MS;
   AryTypePara[273].Other."String" := '';
   AryTypePara[274].TypeName := '';
   AryTypePara[274].bit.Bit0 := FALSE;
   AryTypePara[274].bit.sp := 16#0000;
   AryTypePara[274].bit.Other.Bool_1 := FALSE;
   AryTypePara[274].bit.Other.Byte_2 := 16#00;
   AryTypePara[274].bit.Other.Int_1 := 0;
   AryTypePara[274].bit.Other."Char" := ' ';
   AryTypePara[274].Other.STxxxCCDProgNO := 0;
   AryTypePara[274].Other.FixtureEnable := FALSE;
   AryTypePara[274].Other.Byte_1 := 16#00;
   AryTypePara[274].Other.Int_1 := 0;
   AryTypePara[274].Other."Char" := ' ';
   AryTypePara[274].Other.Word_1 := 16#0000;
   AryTypePara[274].Other.DInt_1 := 0;
   AryTypePara[274].Other.DWord_1 := 16#0000_0000;
   AryTypePara[274].Other.Real_1 := 0.0;
   AryTypePara[274].Other.S5Time := T#0MS;
   AryTypePara[274].Other."String" := '';
   AryTypePara[275].TypeName := '';
   AryTypePara[275].bit.Bit0 := FALSE;
   AryTypePara[275].bit.sp := 16#0000;
   AryTypePara[275].bit.Other.Bool_1 := FALSE;
   AryTypePara[275].bit.Other.Byte_2 := 16#00;
   AryTypePara[275].bit.Other.Int_1 := 0;
   AryTypePara[275].bit.Other."Char" := ' ';
   AryTypePara[275].Other.STxxxCCDProgNO := 0;
   AryTypePara[275].Other.FixtureEnable := FALSE;
   AryTypePara[275].Other.Byte_1 := 16#00;
   AryTypePara[275].Other.Int_1 := 0;
   AryTypePara[275].Other."Char" := ' ';
   AryTypePara[275].Other.Word_1 := 16#0000;
   AryTypePara[275].Other.DInt_1 := 0;
   AryTypePara[275].Other.DWord_1 := 16#0000_0000;
   AryTypePara[275].Other.Real_1 := 0.0;
   AryTypePara[275].Other.S5Time := T#0MS;
   AryTypePara[275].Other."String" := '';
   AryTypePara[276].TypeName := '';
   AryTypePara[276].bit.Bit0 := FALSE;
   AryTypePara[276].bit.sp := 16#0000;
   AryTypePara[276].bit.Other.Bool_1 := FALSE;
   AryTypePara[276].bit.Other.Byte_2 := 16#00;
   AryTypePara[276].bit.Other.Int_1 := 0;
   AryTypePara[276].bit.Other."Char" := ' ';
   AryTypePara[276].Other.STxxxCCDProgNO := 0;
   AryTypePara[276].Other.FixtureEnable := FALSE;
   AryTypePara[276].Other.Byte_1 := 16#00;
   AryTypePara[276].Other.Int_1 := 0;
   AryTypePara[276].Other."Char" := ' ';
   AryTypePara[276].Other.Word_1 := 16#0000;
   AryTypePara[276].Other.DInt_1 := 0;
   AryTypePara[276].Other.DWord_1 := 16#0000_0000;
   AryTypePara[276].Other.Real_1 := 0.0;
   AryTypePara[276].Other.S5Time := T#0MS;
   AryTypePara[276].Other."String" := '';
   AryTypePara[277].TypeName := '';
   AryTypePara[277].bit.Bit0 := FALSE;
   AryTypePara[277].bit.sp := 16#0000;
   AryTypePara[277].bit.Other.Bool_1 := FALSE;
   AryTypePara[277].bit.Other.Byte_2 := 16#00;
   AryTypePara[277].bit.Other.Int_1 := 0;
   AryTypePara[277].bit.Other."Char" := ' ';
   AryTypePara[277].Other.STxxxCCDProgNO := 0;
   AryTypePara[277].Other.FixtureEnable := FALSE;
   AryTypePara[277].Other.Byte_1 := 16#00;
   AryTypePara[277].Other.Int_1 := 0;
   AryTypePara[277].Other."Char" := ' ';
   AryTypePara[277].Other.Word_1 := 16#0000;
   AryTypePara[277].Other.DInt_1 := 0;
   AryTypePara[277].Other.DWord_1 := 16#0000_0000;
   AryTypePara[277].Other.Real_1 := 0.0;
   AryTypePara[277].Other.S5Time := T#0MS;
   AryTypePara[277].Other."String" := '';
   AryTypePara[278].TypeName := '';
   AryTypePara[278].bit.Bit0 := FALSE;
   AryTypePara[278].bit.sp := 16#0000;
   AryTypePara[278].bit.Other.Bool_1 := FALSE;
   AryTypePara[278].bit.Other.Byte_2 := 16#00;
   AryTypePara[278].bit.Other.Int_1 := 0;
   AryTypePara[278].bit.Other."Char" := ' ';
   AryTypePara[278].Other.STxxxCCDProgNO := 0;
   AryTypePara[278].Other.FixtureEnable := FALSE;
   AryTypePara[278].Other.Byte_1 := 16#00;
   AryTypePara[278].Other.Int_1 := 0;
   AryTypePara[278].Other."Char" := ' ';
   AryTypePara[278].Other.Word_1 := 16#0000;
   AryTypePara[278].Other.DInt_1 := 0;
   AryTypePara[278].Other.DWord_1 := 16#0000_0000;
   AryTypePara[278].Other.Real_1 := 0.0;
   AryTypePara[278].Other.S5Time := T#0MS;
   AryTypePara[278].Other."String" := '';
   AryTypePara[279].TypeName := '';
   AryTypePara[279].bit.Bit0 := FALSE;
   AryTypePara[279].bit.sp := 16#0000;
   AryTypePara[279].bit.Other.Bool_1 := FALSE;
   AryTypePara[279].bit.Other.Byte_2 := 16#00;
   AryTypePara[279].bit.Other.Int_1 := 0;
   AryTypePara[279].bit.Other."Char" := ' ';
   AryTypePara[279].Other.STxxxCCDProgNO := 0;
   AryTypePara[279].Other.FixtureEnable := FALSE;
   AryTypePara[279].Other.Byte_1 := 16#00;
   AryTypePara[279].Other.Int_1 := 0;
   AryTypePara[279].Other."Char" := ' ';
   AryTypePara[279].Other.Word_1 := 16#0000;
   AryTypePara[279].Other.DInt_1 := 0;
   AryTypePara[279].Other.DWord_1 := 16#0000_0000;
   AryTypePara[279].Other.Real_1 := 0.0;
   AryTypePara[279].Other.S5Time := T#0MS;
   AryTypePara[279].Other."String" := '';
   AryTypePara[280].TypeName := '';
   AryTypePara[280].bit.Bit0 := FALSE;
   AryTypePara[280].bit.sp := 16#0000;
   AryTypePara[280].bit.Other.Bool_1 := FALSE;
   AryTypePara[280].bit.Other.Byte_2 := 16#00;
   AryTypePara[280].bit.Other.Int_1 := 0;
   AryTypePara[280].bit.Other."Char" := ' ';
   AryTypePara[280].Other.STxxxCCDProgNO := 0;
   AryTypePara[280].Other.FixtureEnable := FALSE;
   AryTypePara[280].Other.Byte_1 := 16#00;
   AryTypePara[280].Other.Int_1 := 0;
   AryTypePara[280].Other."Char" := ' ';
   AryTypePara[280].Other.Word_1 := 16#0000;
   AryTypePara[280].Other.DInt_1 := 0;
   AryTypePara[280].Other.DWord_1 := 16#0000_0000;
   AryTypePara[280].Other.Real_1 := 0.0;
   AryTypePara[280].Other.S5Time := T#0MS;
   AryTypePara[280].Other."String" := '';
   AryTypePara[281].TypeName := '';
   AryTypePara[281].bit.Bit0 := FALSE;
   AryTypePara[281].bit.sp := 16#0000;
   AryTypePara[281].bit.Other.Bool_1 := FALSE;
   AryTypePara[281].bit.Other.Byte_2 := 16#00;
   AryTypePara[281].bit.Other.Int_1 := 0;
   AryTypePara[281].bit.Other."Char" := ' ';
   AryTypePara[281].Other.STxxxCCDProgNO := 0;
   AryTypePara[281].Other.FixtureEnable := FALSE;
   AryTypePara[281].Other.Byte_1 := 16#00;
   AryTypePara[281].Other.Int_1 := 0;
   AryTypePara[281].Other."Char" := ' ';
   AryTypePara[281].Other.Word_1 := 16#0000;
   AryTypePara[281].Other.DInt_1 := 0;
   AryTypePara[281].Other.DWord_1 := 16#0000_0000;
   AryTypePara[281].Other.Real_1 := 0.0;
   AryTypePara[281].Other.S5Time := T#0MS;
   AryTypePara[281].Other."String" := '';
   AryTypePara[282].TypeName := '';
   AryTypePara[282].bit.Bit0 := FALSE;
   AryTypePara[282].bit.sp := 16#0000;
   AryTypePara[282].bit.Other.Bool_1 := FALSE;
   AryTypePara[282].bit.Other.Byte_2 := 16#00;
   AryTypePara[282].bit.Other.Int_1 := 0;
   AryTypePara[282].bit.Other."Char" := ' ';
   AryTypePara[282].Other.STxxxCCDProgNO := 0;
   AryTypePara[282].Other.FixtureEnable := FALSE;
   AryTypePara[282].Other.Byte_1 := 16#00;
   AryTypePara[282].Other.Int_1 := 0;
   AryTypePara[282].Other."Char" := ' ';
   AryTypePara[282].Other.Word_1 := 16#0000;
   AryTypePara[282].Other.DInt_1 := 0;
   AryTypePara[282].Other.DWord_1 := 16#0000_0000;
   AryTypePara[282].Other.Real_1 := 0.0;
   AryTypePara[282].Other.S5Time := T#0MS;
   AryTypePara[282].Other."String" := '';
   AryTypePara[283].TypeName := '';
   AryTypePara[283].bit.Bit0 := FALSE;
   AryTypePara[283].bit.sp := 16#0000;
   AryTypePara[283].bit.Other.Bool_1 := FALSE;
   AryTypePara[283].bit.Other.Byte_2 := 16#00;
   AryTypePara[283].bit.Other.Int_1 := 0;
   AryTypePara[283].bit.Other."Char" := ' ';
   AryTypePara[283].Other.STxxxCCDProgNO := 0;
   AryTypePara[283].Other.FixtureEnable := FALSE;
   AryTypePara[283].Other.Byte_1 := 16#00;
   AryTypePara[283].Other.Int_1 := 0;
   AryTypePara[283].Other."Char" := ' ';
   AryTypePara[283].Other.Word_1 := 16#0000;
   AryTypePara[283].Other.DInt_1 := 0;
   AryTypePara[283].Other.DWord_1 := 16#0000_0000;
   AryTypePara[283].Other.Real_1 := 0.0;
   AryTypePara[283].Other.S5Time := T#0MS;
   AryTypePara[283].Other."String" := '';
   AryTypePara[284].TypeName := '';
   AryTypePara[284].bit.Bit0 := FALSE;
   AryTypePara[284].bit.sp := 16#0000;
   AryTypePara[284].bit.Other.Bool_1 := FALSE;
   AryTypePara[284].bit.Other.Byte_2 := 16#00;
   AryTypePara[284].bit.Other.Int_1 := 0;
   AryTypePara[284].bit.Other."Char" := ' ';
   AryTypePara[284].Other.STxxxCCDProgNO := 0;
   AryTypePara[284].Other.FixtureEnable := FALSE;
   AryTypePara[284].Other.Byte_1 := 16#00;
   AryTypePara[284].Other.Int_1 := 0;
   AryTypePara[284].Other."Char" := ' ';
   AryTypePara[284].Other.Word_1 := 16#0000;
   AryTypePara[284].Other.DInt_1 := 0;
   AryTypePara[284].Other.DWord_1 := 16#0000_0000;
   AryTypePara[284].Other.Real_1 := 0.0;
   AryTypePara[284].Other.S5Time := T#0MS;
   AryTypePara[284].Other."String" := '';
   AryTypePara[285].TypeName := '';
   AryTypePara[285].bit.Bit0 := FALSE;
   AryTypePara[285].bit.sp := 16#0000;
   AryTypePara[285].bit.Other.Bool_1 := FALSE;
   AryTypePara[285].bit.Other.Byte_2 := 16#00;
   AryTypePara[285].bit.Other.Int_1 := 0;
   AryTypePara[285].bit.Other."Char" := ' ';
   AryTypePara[285].Other.STxxxCCDProgNO := 0;
   AryTypePara[285].Other.FixtureEnable := FALSE;
   AryTypePara[285].Other.Byte_1 := 16#00;
   AryTypePara[285].Other.Int_1 := 0;
   AryTypePara[285].Other."Char" := ' ';
   AryTypePara[285].Other.Word_1 := 16#0000;
   AryTypePara[285].Other.DInt_1 := 0;
   AryTypePara[285].Other.DWord_1 := 16#0000_0000;
   AryTypePara[285].Other.Real_1 := 0.0;
   AryTypePara[285].Other.S5Time := T#0MS;
   AryTypePara[285].Other."String" := '';
   AryTypePara[286].TypeName := '';
   AryTypePara[286].bit.Bit0 := FALSE;
   AryTypePara[286].bit.sp := 16#0000;
   AryTypePara[286].bit.Other.Bool_1 := FALSE;
   AryTypePara[286].bit.Other.Byte_2 := 16#00;
   AryTypePara[286].bit.Other.Int_1 := 0;
   AryTypePara[286].bit.Other."Char" := ' ';
   AryTypePara[286].Other.STxxxCCDProgNO := 0;
   AryTypePara[286].Other.FixtureEnable := FALSE;
   AryTypePara[286].Other.Byte_1 := 16#00;
   AryTypePara[286].Other.Int_1 := 0;
   AryTypePara[286].Other."Char" := ' ';
   AryTypePara[286].Other.Word_1 := 16#0000;
   AryTypePara[286].Other.DInt_1 := 0;
   AryTypePara[286].Other.DWord_1 := 16#0000_0000;
   AryTypePara[286].Other.Real_1 := 0.0;
   AryTypePara[286].Other.S5Time := T#0MS;
   AryTypePara[286].Other."String" := '';
   AryTypePara[287].TypeName := '';
   AryTypePara[287].bit.Bit0 := FALSE;
   AryTypePara[287].bit.sp := 16#0000;
   AryTypePara[287].bit.Other.Bool_1 := FALSE;
   AryTypePara[287].bit.Other.Byte_2 := 16#00;
   AryTypePara[287].bit.Other.Int_1 := 0;
   AryTypePara[287].bit.Other."Char" := ' ';
   AryTypePara[287].Other.STxxxCCDProgNO := 0;
   AryTypePara[287].Other.FixtureEnable := FALSE;
   AryTypePara[287].Other.Byte_1 := 16#00;
   AryTypePara[287].Other.Int_1 := 0;
   AryTypePara[287].Other."Char" := ' ';
   AryTypePara[287].Other.Word_1 := 16#0000;
   AryTypePara[287].Other.DInt_1 := 0;
   AryTypePara[287].Other.DWord_1 := 16#0000_0000;
   AryTypePara[287].Other.Real_1 := 0.0;
   AryTypePara[287].Other.S5Time := T#0MS;
   AryTypePara[287].Other."String" := '';
   AryTypePara[288].TypeName := '';
   AryTypePara[288].bit.Bit0 := FALSE;
   AryTypePara[288].bit.sp := 16#0000;
   AryTypePara[288].bit.Other.Bool_1 := FALSE;
   AryTypePara[288].bit.Other.Byte_2 := 16#00;
   AryTypePara[288].bit.Other.Int_1 := 0;
   AryTypePara[288].bit.Other."Char" := ' ';
   AryTypePara[288].Other.STxxxCCDProgNO := 0;
   AryTypePara[288].Other.FixtureEnable := FALSE;
   AryTypePara[288].Other.Byte_1 := 16#00;
   AryTypePara[288].Other.Int_1 := 0;
   AryTypePara[288].Other."Char" := ' ';
   AryTypePara[288].Other.Word_1 := 16#0000;
   AryTypePara[288].Other.DInt_1 := 0;
   AryTypePara[288].Other.DWord_1 := 16#0000_0000;
   AryTypePara[288].Other.Real_1 := 0.0;
   AryTypePara[288].Other.S5Time := T#0MS;
   AryTypePara[288].Other."String" := '';
   AryTypePara[289].TypeName := '';
   AryTypePara[289].bit.Bit0 := FALSE;
   AryTypePara[289].bit.sp := 16#0000;
   AryTypePara[289].bit.Other.Bool_1 := FALSE;
   AryTypePara[289].bit.Other.Byte_2 := 16#00;
   AryTypePara[289].bit.Other.Int_1 := 0;
   AryTypePara[289].bit.Other."Char" := ' ';
   AryTypePara[289].Other.STxxxCCDProgNO := 0;
   AryTypePara[289].Other.FixtureEnable := FALSE;
   AryTypePara[289].Other.Byte_1 := 16#00;
   AryTypePara[289].Other.Int_1 := 0;
   AryTypePara[289].Other."Char" := ' ';
   AryTypePara[289].Other.Word_1 := 16#0000;
   AryTypePara[289].Other.DInt_1 := 0;
   AryTypePara[289].Other.DWord_1 := 16#0000_0000;
   AryTypePara[289].Other.Real_1 := 0.0;
   AryTypePara[289].Other.S5Time := T#0MS;
   AryTypePara[289].Other."String" := '';
   AryTypePara[290].TypeName := '';
   AryTypePara[290].bit.Bit0 := FALSE;
   AryTypePara[290].bit.sp := 16#0000;
   AryTypePara[290].bit.Other.Bool_1 := FALSE;
   AryTypePara[290].bit.Other.Byte_2 := 16#00;
   AryTypePara[290].bit.Other.Int_1 := 0;
   AryTypePara[290].bit.Other."Char" := ' ';
   AryTypePara[290].Other.STxxxCCDProgNO := 0;
   AryTypePara[290].Other.FixtureEnable := FALSE;
   AryTypePara[290].Other.Byte_1 := 16#00;
   AryTypePara[290].Other.Int_1 := 0;
   AryTypePara[290].Other."Char" := ' ';
   AryTypePara[290].Other.Word_1 := 16#0000;
   AryTypePara[290].Other.DInt_1 := 0;
   AryTypePara[290].Other.DWord_1 := 16#0000_0000;
   AryTypePara[290].Other.Real_1 := 0.0;
   AryTypePara[290].Other.S5Time := T#0MS;
   AryTypePara[290].Other."String" := '';
   AryTypePara[291].TypeName := '';
   AryTypePara[291].bit.Bit0 := FALSE;
   AryTypePara[291].bit.sp := 16#0000;
   AryTypePara[291].bit.Other.Bool_1 := FALSE;
   AryTypePara[291].bit.Other.Byte_2 := 16#00;
   AryTypePara[291].bit.Other.Int_1 := 0;
   AryTypePara[291].bit.Other."Char" := ' ';
   AryTypePara[291].Other.STxxxCCDProgNO := 0;
   AryTypePara[291].Other.FixtureEnable := FALSE;
   AryTypePara[291].Other.Byte_1 := 16#00;
   AryTypePara[291].Other.Int_1 := 0;
   AryTypePara[291].Other."Char" := ' ';
   AryTypePara[291].Other.Word_1 := 16#0000;
   AryTypePara[291].Other.DInt_1 := 0;
   AryTypePara[291].Other.DWord_1 := 16#0000_0000;
   AryTypePara[291].Other.Real_1 := 0.0;
   AryTypePara[291].Other.S5Time := T#0MS;
   AryTypePara[291].Other."String" := '';
   AryTypePara[292].TypeName := '';
   AryTypePara[292].bit.Bit0 := FALSE;
   AryTypePara[292].bit.sp := 16#0000;
   AryTypePara[292].bit.Other.Bool_1 := FALSE;
   AryTypePara[292].bit.Other.Byte_2 := 16#00;
   AryTypePara[292].bit.Other.Int_1 := 0;
   AryTypePara[292].bit.Other."Char" := ' ';
   AryTypePara[292].Other.STxxxCCDProgNO := 0;
   AryTypePara[292].Other.FixtureEnable := FALSE;
   AryTypePara[292].Other.Byte_1 := 16#00;
   AryTypePara[292].Other.Int_1 := 0;
   AryTypePara[292].Other."Char" := ' ';
   AryTypePara[292].Other.Word_1 := 16#0000;
   AryTypePara[292].Other.DInt_1 := 0;
   AryTypePara[292].Other.DWord_1 := 16#0000_0000;
   AryTypePara[292].Other.Real_1 := 0.0;
   AryTypePara[292].Other.S5Time := T#0MS;
   AryTypePara[292].Other."String" := '';
   AryTypePara[293].TypeName := '';
   AryTypePara[293].bit.Bit0 := FALSE;
   AryTypePara[293].bit.sp := 16#0000;
   AryTypePara[293].bit.Other.Bool_1 := FALSE;
   AryTypePara[293].bit.Other.Byte_2 := 16#00;
   AryTypePara[293].bit.Other.Int_1 := 0;
   AryTypePara[293].bit.Other."Char" := ' ';
   AryTypePara[293].Other.STxxxCCDProgNO := 0;
   AryTypePara[293].Other.FixtureEnable := FALSE;
   AryTypePara[293].Other.Byte_1 := 16#00;
   AryTypePara[293].Other.Int_1 := 0;
   AryTypePara[293].Other."Char" := ' ';
   AryTypePara[293].Other.Word_1 := 16#0000;
   AryTypePara[293].Other.DInt_1 := 0;
   AryTypePara[293].Other.DWord_1 := 16#0000_0000;
   AryTypePara[293].Other.Real_1 := 0.0;
   AryTypePara[293].Other.S5Time := T#0MS;
   AryTypePara[293].Other."String" := '';
   AryTypePara[294].TypeName := '';
   AryTypePara[294].bit.Bit0 := FALSE;
   AryTypePara[294].bit.sp := 16#0000;
   AryTypePara[294].bit.Other.Bool_1 := FALSE;
   AryTypePara[294].bit.Other.Byte_2 := 16#00;
   AryTypePara[294].bit.Other.Int_1 := 0;
   AryTypePara[294].bit.Other."Char" := ' ';
   AryTypePara[294].Other.STxxxCCDProgNO := 0;
   AryTypePara[294].Other.FixtureEnable := FALSE;
   AryTypePara[294].Other.Byte_1 := 16#00;
   AryTypePara[294].Other.Int_1 := 0;
   AryTypePara[294].Other."Char" := ' ';
   AryTypePara[294].Other.Word_1 := 16#0000;
   AryTypePara[294].Other.DInt_1 := 0;
   AryTypePara[294].Other.DWord_1 := 16#0000_0000;
   AryTypePara[294].Other.Real_1 := 0.0;
   AryTypePara[294].Other.S5Time := T#0MS;
   AryTypePara[294].Other."String" := '';
   AryTypePara[295].TypeName := '';
   AryTypePara[295].bit.Bit0 := FALSE;
   AryTypePara[295].bit.sp := 16#0000;
   AryTypePara[295].bit.Other.Bool_1 := FALSE;
   AryTypePara[295].bit.Other.Byte_2 := 16#00;
   AryTypePara[295].bit.Other.Int_1 := 0;
   AryTypePara[295].bit.Other."Char" := ' ';
   AryTypePara[295].Other.STxxxCCDProgNO := 0;
   AryTypePara[295].Other.FixtureEnable := FALSE;
   AryTypePara[295].Other.Byte_1 := 16#00;
   AryTypePara[295].Other.Int_1 := 0;
   AryTypePara[295].Other."Char" := ' ';
   AryTypePara[295].Other.Word_1 := 16#0000;
   AryTypePara[295].Other.DInt_1 := 0;
   AryTypePara[295].Other.DWord_1 := 16#0000_0000;
   AryTypePara[295].Other.Real_1 := 0.0;
   AryTypePara[295].Other.S5Time := T#0MS;
   AryTypePara[295].Other."String" := '';
   AryTypePara[296].TypeName := '';
   AryTypePara[296].bit.Bit0 := FALSE;
   AryTypePara[296].bit.sp := 16#0000;
   AryTypePara[296].bit.Other.Bool_1 := FALSE;
   AryTypePara[296].bit.Other.Byte_2 := 16#00;
   AryTypePara[296].bit.Other.Int_1 := 0;
   AryTypePara[296].bit.Other."Char" := ' ';
   AryTypePara[296].Other.STxxxCCDProgNO := 0;
   AryTypePara[296].Other.FixtureEnable := FALSE;
   AryTypePara[296].Other.Byte_1 := 16#00;
   AryTypePara[296].Other.Int_1 := 0;
   AryTypePara[296].Other."Char" := ' ';
   AryTypePara[296].Other.Word_1 := 16#0000;
   AryTypePara[296].Other.DInt_1 := 0;
   AryTypePara[296].Other.DWord_1 := 16#0000_0000;
   AryTypePara[296].Other.Real_1 := 0.0;
   AryTypePara[296].Other.S5Time := T#0MS;
   AryTypePara[296].Other."String" := '';
   AryTypePara[297].TypeName := '';
   AryTypePara[297].bit.Bit0 := FALSE;
   AryTypePara[297].bit.sp := 16#0000;
   AryTypePara[297].bit.Other.Bool_1 := FALSE;
   AryTypePara[297].bit.Other.Byte_2 := 16#00;
   AryTypePara[297].bit.Other.Int_1 := 0;
   AryTypePara[297].bit.Other."Char" := ' ';
   AryTypePara[297].Other.STxxxCCDProgNO := 0;
   AryTypePara[297].Other.FixtureEnable := FALSE;
   AryTypePara[297].Other.Byte_1 := 16#00;
   AryTypePara[297].Other.Int_1 := 0;
   AryTypePara[297].Other."Char" := ' ';
   AryTypePara[297].Other.Word_1 := 16#0000;
   AryTypePara[297].Other.DInt_1 := 0;
   AryTypePara[297].Other.DWord_1 := 16#0000_0000;
   AryTypePara[297].Other.Real_1 := 0.0;
   AryTypePara[297].Other.S5Time := T#0MS;
   AryTypePara[297].Other."String" := '';
   AryTypePara[298].bit.Bit0 := FALSE;
   AryTypePara[298].bit.sp := 16#0000;
   AryTypePara[298].bit.Other.Bool_1 := FALSE;
   AryTypePara[298].bit.Other.Byte_2 := 16#00;
   AryTypePara[298].bit.Other.Int_1 := 0;
   AryTypePara[298].bit.Other."Char" := ' ';
   AryTypePara[298].Other.FixtureEnable := FALSE;
   AryTypePara[298].Other.Byte_1 := 16#00;
   AryTypePara[298].Other.Int_1 := 0;
   AryTypePara[298].Other."Char" := ' ';
   AryTypePara[298].Other.Word_1 := 16#0000;
   AryTypePara[298].Other.DInt_1 := 0;
   AryTypePara[298].Other.DWord_1 := 16#0000_0000;
   AryTypePara[298].Other.Real_1 := 0.0;
   AryTypePara[298].Other.S5Time := T#0MS;
   AryTypePara[298].Other."String" := '';
   AryTypePara[299].bit.Bit0 := FALSE;
   AryTypePara[299].bit.sp := 16#0000;
   AryTypePara[299].bit.Other.Bool_1 := FALSE;
   AryTypePara[299].bit.Other.Byte_2 := 16#00;
   AryTypePara[299].bit.Other.Int_1 := 0;
   AryTypePara[299].bit.Other."Char" := ' ';
   AryTypePara[299].Other.FixtureEnable := FALSE;
   AryTypePara[299].Other.Byte_1 := 16#00;
   AryTypePara[299].Other.Int_1 := 0;
   AryTypePara[299].Other."Char" := ' ';
   AryTypePara[299].Other.Word_1 := 16#0000;
   AryTypePara[299].Other.DInt_1 := 0;
   AryTypePara[299].Other.DWord_1 := 16#0000_0000;
   AryTypePara[299].Other.Real_1 := 0.0;
   AryTypePara[299].Other.S5Time := T#0MS;
   AryTypePara[299].Other."String" := '';
   AryTypePara[300].bit.Bit0 := FALSE;
   AryTypePara[300].bit.sp := 16#0000;
   AryTypePara[300].bit.Other.Bool_1 := FALSE;
   AryTypePara[300].bit.Other.Byte_2 := 16#00;
   AryTypePara[300].bit.Other.Int_1 := 0;
   AryTypePara[300].bit.Other."Char" := ' ';
   AryTypePara[300].Other.FixtureEnable := FALSE;
   AryTypePara[300].Other.Byte_1 := 16#00;
   AryTypePara[300].Other.Int_1 := 0;
   AryTypePara[300].Other."Char" := ' ';
   AryTypePara[300].Other.Word_1 := 16#0000;
   AryTypePara[300].Other.DInt_1 := 0;
   AryTypePara[300].Other.DWord_1 := 16#0000_0000;
   AryTypePara[300].Other.Real_1 := 0.0;
   AryTypePara[300].Other.S5Time := T#0MS;
   AryTypePara[300].Other."String" := '';
END_DATA_BLOCK

// folder: 001_KL_Standard_FB

DATA_BLOCK "DB1000_StdSignal"   // DB1000
{ S7_Optimized_Access := 'TRUE' }
VERSION : 0.0
// stored: InstanceOfName FB1000_StdSignal
"FB1000_StdSignal"
BEGIN
END_DATA_BLOCK

DATA_BLOCK "DB1009_Constant"   // DB1009
{ S7_Optimized_Access := 'FALSE' }
VERSION : 0.1
   VAR
      ConnectID : Struct   // TCP连接ID
         ID101 : Int := 101;
         ID102 : Int := 102;
         ID103 : Int := 103;
         ID104 : Int := 104;
         ID105 : Int := 105;
         ID106 : Int := 106;
         ID107 : Int := 107;
         ID108 : Int := 108;
         ID109 : Int := 109;
         ID110 : Int := 110;
         ID111 : Int := 111;
         ID112 : Int := 112;
         ID113 : Int := 113;
         ID114 : Int := 114;
         ID115 : Int := 115;
         ID116 : Int := 116;
         ID117 : Int := 117;
         ID118 : Int := 118;
         ID119 : Int := 119;
         ID120 : Int := 119;
      END_STRUCT;
      falseBool : Bool;
      trueBool : Bool;
      EmptyByte : Byte;
      EmptyInt : Int;
      EmptyDint : DInt;
      EmptyStr : String[1];
      KeyenceCodeReaderSend : String[3] := 'LON';
      KeyenceCodeReaderErr : String[5] := 'ERROR';
   END_VAR
BEGIN
END_DATA_BLOCK

DATA_BLOCK "DB1200_FB_std_Switch"   // DB1200
{ S7_Optimized_Access := 'TRUE' }
VERSION : 0.1
// stored: InstanceOfName FB1200_std_Switch
"FB1200_std_Switch"
BEGIN
END_DATA_BLOCK

DATA_BLOCK "DB1202_IOCheck"   // DB1202
{ S7_Optimized_Access := 'TRUE' }
VERSION : 0.1
// stored: InstanceOfName FB1202_IOCheck_
"FB1202_IOCheck_"
BEGIN
END_DATA_BLOCK

DATA_BLOCK "DB1210_DPRD_DPWR"   // DB1210
{ S7_Optimized_Access := 'TRUE' }
VERSION : 0.1
// stored: InstanceOfName FB1210_DPRD_DPWR
"FB1210_DPRD_DPWR"
BEGIN
END_DATA_BLOCK

// folder: 002_Err_Prompt_Handle

DATA_BLOCK "DB1140_Message"   // DB1140
{ S7_Optimized_Access := 'TRUE' }
VERSION : 0.1
// stored: InstanceOfName FB1140_Message
"FB1140_Message"
BEGIN
END_DATA_BLOCK

DATA_BLOCK "DB1142_TypeChangePrompt"   // DB1142
{ S7_Optimized_Access := 'TRUE' }
VERSION : 0.1
// stored: InstanceOfName FB1142_TypeChangePrompt
"FB1142_TypeChangePrompt"
BEGIN
END_DATA_BLOCK

DATA_BLOCK "DB1146_PromptFree"   // DB1146
{ S7_Optimized_Access := 'FALSE' }
VERSION : 0.1
   VAR
      Public : Struct
         OperationNotPmt : Bool;   // 气缸操作被禁止，请检查安全条件！
         StepMode : Bool;   // 设备处于单步模式，请注意安全！
         EmptyMode : Bool;   // 设备已经开始清空，请等待！
         AutoModeOffPrompt : Bool;   // 等待循环结束，暂停自动模式中！
         DoorOveRideStarting : Bool;   // 开始安全门旁路,等待各流程结束!
         OkToStart : Bool;   // 请启动设备！
         WaitPcCommond : Bool;   // 等待PC命令！
         LightCurtain : Bool;   // 光幕被遮,注意安全!
         AutoModeNotStarted : Bool;   // 请摁下自动模式启动按钮！
         AskPcData : Bool;   // 请求上位机参数录入...
         PleaseChangeTool : Bool;   // 请开始换夹具...
         AskPcData_1 : Bool;   // 请求上位机参数录入...
         do_ChgGrp_Act : Bool;   // 换爪运行中
         do_HorDril_Act : Bool;   // 水平方向钻入运行中
         do_UpDril_Act : Bool;   // 向上方向钻入运行中
         do_DownDril_Act : Bool;   // 向下方向钻入运行中
         do_ChkScrew_Act : Bool;   // 检查钻头运行中
         do_Clean_Act : Bool;   // 清洁运行中
         do_ChgGrp_Pos : Bool;   // 换爪位置
         do_HorDril_Pos : Bool;   // 水平方向钻入位置
         do_UpDril_Pos : Bool;   // 向上方向钻入位置
         do_DownDril_Pos : Bool;   // 向下方向钻入位置
         do_ChkScrew_Pos : Bool;   // 检查钻头位置
         do_ReqDrilling : Bool;   // 请求钻孔
         do_ReqStopDril : Bool;   // 请求停止钻孔
         do_Clean_Pos : Bool;   // 清洁位置
         do_ChgGrp_Don : Bool;   // 换爪完成
         do_HorDril_Don : Bool;   // 水平方向钻入完成
         do_UpDril_Don : Bool;   // 向上方向钻入完成
         do_DownDril_Don : Bool;   // 向下方向钻入完成
         do_ChkScrew_Don : Bool;   // 检查钻头完成
      END_STRUCT;
      ST01 : Struct
         Z01ExtIng : Bool;   // Z01.解锁缸到工作位置...
         Z01RetIng : Bool;   // Z01.解锁缸到基本位置...
         Z02ExtIng : Bool;   // Z02.备用到工作位置...
         Z02RetIng : Bool;   // Z02.备用到基本位置...
         Z03ExtIng : Bool;   // Z03.备用到工作位置...
         Z03RetIng : Bool;   // Z03.备用到基本位置...
         Z04ExtIng : Bool;   // Z04.备用到工作位置...
         Z04RetIng : Bool;   // Z04.备用到基本位置...
         Z05ExtIng : Bool;   // Z05.备用到工作位置...
         Z05RetIng : Bool;   // Z05.备用到基本位置...
         Z06Exting : Bool;
         Z06Reting : Bool;
         Z07Exting : Bool;
         Z07Reting : Bool;
         Z08Exting : Bool;
         Z08Reting : Bool;
         Z09Exting : Bool;
         Z09Reting : Bool;
         Z10Exting : Bool;
         Z10Reting : Bool;
         WaitZ01Ext_0 : Bool;   // 等待推力缸完全释放
         WaitZ01Ext_1 : Bool;   // 等待推力缸完全释放
         WaitZ01Ext_2 : Bool;   // 等待推力缸完全释放
         Z11Exting : Bool;
         Z11Reting : Bool;
         HeatMachin : Bool;   // 热机中...
         Spare7_2 : Bool;
         Spare7_3 : Bool;
         Spare7_4 : Bool;
         Spare7_5 : Bool;
         Spare7_6 : Bool;
         Spare7_7 : Bool;
      END_STRUCT;
   END_VAR
BEGIN
END_DATA_BLOCK

DATA_BLOCK "DB1147_PromptStartNotPmt"   // DB1147
{ S7_Optimized_Access := 'FALSE' }
VERSION : 0.1
   VAR
      Public : Struct
         ToBeHomePos : Bool;   // 设备不在原点,需要复位!
         AutoModeNotStarted : Bool;   // 请摁下自动模式启动按钮！
         DoorOveRideStarted : Bool;   // 安全门旁路，注意安全！
         DoorLockFail : Bool;   // 安全门电磁线圈锁定失败！
         PcCommErr : Bool;   // 上位机通讯失败！
         VisualPCComErr : Bool := false;   // 视觉主机通讯失败！
         ParaWiriteOuttime : Bool;   // 上位机写入参数超时！
         ChangeHorDrillSlab : Bool;   // 水平锤钻水泥板已打完，请更换水泥板！
         ChangeUploadSlab : Bool;   // 垂直向上水泥板已打完，请更换水泥板！
         ChangeDownloadSlab : Bool;   // 垂直向下水泥板已打完，请更换水泥板！
         ChangeHorVChiselSlab : Bool;   // 水平凿击水泥板已打完，请更换水泥板！
         FTComErr : Bool;   // 力控通讯失败
         xx6 : Bool;   // NotPmt_5
         xx7 : Bool;   // NotPmt_6
         xx8 : Bool;   // NotPmt_7
         xx9 : Bool;   // NotPmt_10
         xx10 : Bool;   // NotPmt_11
         xx11 : Bool;   // NotPmt_12
         xx12 : Bool;   // NotPmt_13
         xx13 : Bool;   // NotPmt_14
         xx14 : Bool;   // NotPmt_15
         xx15 : Bool;   // NotPmt_16
         xx16 : Bool;   // NotPmt_17
         xx17 : Bool;   // NotPmt_20
         xx18 : Bool;   // NotPmt_21
         xx19 : Bool;   // NotPmt_22
         xx20 : Bool;   // NotPmt_23
         xx21 : Bool;   // NotPmt_24
         xx22 : Bool;   // NotPmt_25
         xx23 : Bool;   // NotPmt_26
         xx24 : Bool;   // NotPmt_27
         xx25 : Bool;   // NotPmt_30
      END_STRUCT;
   END_VAR
BEGIN
END_DATA_BLOCK

DATA_BLOCK "DB1148_PromptBeeper"   // DB1148
{ S7_Optimized_Access := 'FALSE' }
VERSION : 0.1
   VAR
      Public : Struct
         EMING : Bool;   // 设备紧急停止中,请复位！
         AirPressureLow : Bool;   // 设备气压低，请复位！
         BitStuckErr_Fixture : Bool;   // 夹具卡死，请人工处理!
         CylinderOPerateNotPmt : Bool;   // 气缸操作条件不满足，请检查！
         PcErr : Bool;   // 上位机急停！
         DrillTimeOut : Bool;   // 打孔超时！
         Z01StartPosErr : Bool;   // 推力缸初始位置不正确！
         DownHeightErr : Bool;   // 向下水泥块厚度不在限制范围内(350-450)
         Spare1_0 : Bool;
         RobotNotReady : Bool;   // 机器人未准备好！
         EMOK : Bool;   // 操作盒急停NOK
         RobotEMOK : Bool;   // 机器人急停按钮NOK
         BitStuckErr_HighCurrent : Bool;   // 钻头卡死，高电流报警！
         InsideEMOK : Bool;   // 围栏内侧急停NOK
         InsideEMOK1 : Bool;   // 水泥块击打框架急停NOK
         FixtureAtPosErr : Bool;   // 取夹具时夹具不在位，请检查夹具状态及感应开关
         PowerToolNoCompErr : Bool;   // 电源夹具ID号错误，请检查夹具！
         CurrentLowTimeOut : Bool;   // 低电流工作超时报警！
         CurrentHighTimeOut : Bool;   // 高电流工作超时报警！
         ForceCannotZero : Bool;   // 加载力数据不能为零!
         HorChiselStuckErr : Bool;   // 水平凿击卡死报警
         DownChiselStuckErr : Bool;   // 向下凿击卡死报警
         RetHome_PowerOff : Bool;   // 手动打孔位置回原点电源未正常通电！
         IoToolNoCompErr : Bool;   // 信号夹具ID号错误，请检查夹具！
         RetHome_Z02RetTimeOut : Bool;   // 手动打孔位置回原点气缸回拉不到位！
         ConcreteEnd : Bool;   // 当前水泥块已用完，请更换！
         DiamondCoreNOK : Bool;   // 水钻岩芯未敲击出，请人工处理！
         ScrLenFault : Bool;   // 批头长度错误，请更换！
         AngleErr : Bool;   // 角度设置超限！
         PutGunPosFull : Bool;   // 夹具位置已满，无法换型！
         DrillDepthErr : Bool;   // 钻孔深度超限！
         RobotSpeed : Bool;   // 机器人设置速度不能超过100！
      END_STRUCT;
      ST01 : Struct
         Z01ExtErr : Bool;   // Z01.推力气缸工作位置故障!%Q4.0
         Z01RetErr : Bool;   // Z01.推力气缸基本位置故障!%I3.3%Q4.1
         Z02ExtErr : Bool;   // Z02.辅助气缸工作位置故障!%I3.2%Q4.2
         Z02RetErr : Bool;   // Z02.辅助气缸基本位置故障!%Q4.3
         Z03ExtErr : Bool;   // Z03.左防尘盖夹紧缸工作位置故障!%I2.4%Q4.4
         Z03RetErr : Bool;   // Z03.左防尘盖夹紧缸基本位置故障!%I2.5%Q4.5
         Z04ExtErr : Bool;   // Z04.右防尘盖夹紧缸工作位置故障!%I3.0%Q4.6
         Z04RetErr : Bool;   // Z04.右防尘盖夹紧缸基本位置故障!%I3.1%Q4.7
         Z05ExtErr : Bool;   // Z05.枪电源工作位置故障!%Q5.0
         Z05RetErr : Bool;   // Z05.枪电源基本位置故障!
         Z06ExtErr : Bool;   // Z06.水钻振动锤工作位置故障!%Q5.1
         Z06RetErr : Bool;   // Z06.水钻振动锤基本位置故障!
         Z07ExtErr : Bool;   // Z07.快换盘锁紧工作位置故障!%Q5.6
         Z07RetErr : Bool;   // Z07.快换盘锁紧基本位置故障!%Q5.7
         Z08ExtErr : Bool;   // Z08.参数写入工作位置故障!
         Z08RetErr : Bool;   // Z08.参数写入基本位置故障!
         Z09ExtErr : Bool;   // Z09.三爪卡盘气缸工作位置故障!
         Z09RetErr : Bool;   // Z09.三爪卡盘气缸基本位置故障!
         Spare6_2 : Bool;
         Spare6_3 : Bool;
         Spare6_4 : Bool;
         Spare6_5 : Bool;
         DrillModeErr : Bool;   // 钻孔模式输入有误！
         ToolPosNotOk : Bool;   // 夹具库枪位置不正确！
         PutToolPosNotOk : Bool;   // 夹具未放到位！
         DrillTimeOutZero : Bool;   // 打孔超时时间不能设置为零！
         DrillTimeZero : Bool;   // 打孔时间不能设置为零！
         CurrentTimeZero : Bool;   // 低电流持续时间不能设置为零！
         Spare7_4 : Bool;
         Spare7_5 : Bool;
         Spare7_6 : Bool;
         Spare7_7 : Bool;
      END_STRUCT;
   END_VAR
BEGIN
END_DATA_BLOCK

// folder: 003_HomeStep

DATA_BLOCK "DB1040_HomePos"   // DB1040
{ S7_Optimized_Access := 'TRUE' }
VERSION : 0.1
// stored: InstanceOfName FB1040_HomePos
"FB1040_HomePos"
BEGIN
END_DATA_BLOCK

// folder: 004_AutoStep

DATA_BLOCK "DB720_KuKa_MainCtrl"   // DB720
{ S7_Optimized_Access := 'TRUE' }
VERSION : 0.1
// stored: InstanceOfName FB720_KuKa_MainCtrl
"FB720_KuKa_MainCtrl"
BEGIN
END_DATA_BLOCK

DATA_BLOCK "DB1042_Timer"   // DB1042
{ S7_Optimized_Access := 'FALSE' }
VERSION : 0.1
   VAR
      Communication : Bool;
      DrillMemory : Bool;   // 用作打击记忆，回原点开枪
      HDrillDepth : Bool;   // 钻孔进给记忆
      DDrillDepth : Bool;   // 钻孔进给记忆
      FirstStart : Bool;   // 第一次开始，不以电流为开始方式
      HTimeOutTimesPLS : Bool;
      DTimeOutTimesPLS : Bool;
      HCLowTimeOutTimesPLS : Bool;
      HCHighTimeOutTimesPLS : Bool;
      DCLowTimeOutTimesPLS : Bool;
      DCHighTimeOutTimesPLS : Bool;
      HTimeOutTimes : Int;   // 水平击打超时次数，超过两次报警
      DTimeOutTimes : Int;   // 向下击打超时次数，超过两次报警
      HCLowTimeOutTimes : Int;   // 水平低电流超时次数，超过两次报警
      HCHighTimeOutTimes : Int;   // 水平高电流超时次数，超过两次报警
      DCLowTimeOutTimes : Int;   // 向下低电流超时次数，超过两次报警
      DCHighTimeOutTimes : Int;   // 向下高电流超时次数，超过两次报警
      Force : Real;
      DrillDirectionMemory : Int;   // 上次钻孔记忆
      DrillDirectionCurrent : Int;   // 上次钻孔方向
      ADDTimer_HorDrill : IEC_TIMER;
      ADDTimer_DownDrill : IEC_TIMER;
      Z02ExtPos : IEC_TIMER;
      Z02ExtPos_1 : IEC_TIMER;
      FirstStartTime : IEC_TIMER;
      HDrillEndTime : IEC_TIMER;
      DDrillEndTime : IEC_TIMER;
      HCurrentLastTime : IEC_TIMER;   // 水平有效电流持续时间
      DCurrentLastTime : IEC_TIMER;   // 向下有效电流持续时间
      CurrentLowTimeOut : IEC_TIMER;   // 低电流超时时间
      CurrentHighTimeOut : IEC_TIMER;   // 高电流超时时间
      GougeTimeOut : IEC_TIMER;   // 凿击超时时间
      GougeTimeOut_1 : IEC_TIMER;   // 斜凿击超时时间
      GougeTimeOut_2 : IEC_TIMER;
      HorChiselTimeOut : IEC_TIMER;   // 水平凿击结束超时
      FixtureStuckTimeOut : IEC_TIMER;   // 夹具卡死超时
      PowerOn_RetHome : IEC_TIMER;
      RetHomeHighCurrentOut : IEC_TIMER;
      RetHome_Z02TimeOut : IEC_TIMER;   // 回原点气缸回拉不到位
      DrillingHighCurrentOut : IEC_TIMER;   // 打孔过程中高电流超时报警
   END_VAR
BEGIN
   // CurrentLowTimeOut.Q : 电流超时时间
   // GougeTimeOut.Q : 凿击超时时间
   // GougeTimeOut_1.Q : 斜凿击超时时间
   // CurrentHighTimeOut.Q : 电流超时时间
   // HCurrentLastTime.Q : 有效电流持续时间
   // DCurrentLastTime.Q : 有效电流持续时间
END_DATA_BLOCK

DATA_BLOCK "DB1060_AutoStep"   // DB1060
{ S7_Optimized_Access := 'FALSE' }
VERSION : 0.1
// stored: InstanceOfName FB1060_AutoStep
"FB1060_AutoStep"
BEGIN
END_DATA_BLOCK

DATA_BLOCK "DB1081_ValveCall"   // DB1081
{ S7_Optimized_Access := 'TRUE' }
VERSION : 0.1
// stored: InstanceOfName FB1081_ValveCall
"FB1081_ValveCall"
BEGIN
END_DATA_BLOCK

DATA_BLOCK "DB1910_DrillData"   // DB1910
{ S7_Optimized_Access := 'TRUE' }
VERSION : 0.1
// stored: InstanceOfName FB1910_DrillData
"FB1910_DrillData"
BEGIN
   HorDrill.SlabLength := 1200.0;
   HorDrill.SlabWidth := 740.0;
   DownDrill.SlabWidth := 1200.0;
   DownDrill.SlabLength := 750.0;
   HorDrill.CurrentDrillWidth := 40.0;
   HorDrill.CurrentDrillLength := 30.0;
   HorDrill.LastDrillWidth := 40.0;
   HorDrill.AlreadyDrillWidth := 485.0;
   HorDrill.AlreadyDrillLength := 990.0;
   HorDrill.MaxWidth := 40.0;
   HorDrill.gi_OffSetY := 1020.0;
   HorDrill.gi_OffSetZ := -485.0;
   HorDrill.PosNo := 35;
   DownDrill.CurrentDrillWidth := 25.0;
   DownDrill.LastDrillWidth := 25.0;
   DownDrill.AlreadyDrillWidth := 175.0;
   DownDrill.MaxWidth := 25.0;
   DownDrill.gi_OffSetY := 1200.0;
   DownDrill.gi_OffSetZ := 200.0;
   DownDrill.PosNo := 1;
   AUX.GougeDrillWidth := 40.0;
END_DATA_BLOCK

// folder: 005_Component

DATA_BLOCK "DB1080_Component"   // DB1080
{ S7_Optimized_Access := 'TRUE' }
VERSION : 0.1
// stored: InstanceOfName FB1080_Component
"FB1080_Component"
BEGIN
END_DATA_BLOCK

DATA_BLOCK "DB1900_Communication_PC"   // DB1900
{ S7_Optimized_Access := 'FALSE' }
VERSION : 0.1
   VAR
      Send : Struct
         Heart : Bool;   // 心跳
         EmmMode : Bool := 0;   // 急停模式
         ManMode : Bool := 0;   // 手动模式
         AutoMode : Bool;   // 自动模式
         PowerOff : Bool := 0;   // 异常停止
         Spare05 : Bool := 0;
         Spare06 : Bool;
         Spare07 : Bool;
         ParaWrite : Bool;   // 请求参数
         DrillStart : Bool;   // 打孔Ready
         DrillRunning : Bool;   // 打孔中
         ChangeToolDone : Bool;   // 收到更换电锤
         WorkDone : Bool;   // 收到作业完成
         WorkStart : Bool;   // 作业开始
         Z01VentValve : Bool;   // 推力气缸中泄
         Z02VentValve : Bool;   // 辅助气缸中泄
         Z01ExtPos : Bool := TRUE;   // 推力气缸伸出
         Z01RetPos : Bool := FALSE;   // 推力气缸缩回
         Z02ExtPos : Bool := FALSE;   // 辅助气缸伸出
         Z02RetPos : Bool := TRUE;   // 辅助气缸缩回
         Z03ExtPos : Bool := FALSE;   // 左防尘盖夹紧缸伸出
         Z03RetPos : Bool := TRUE;   // 左防尘盖夹紧缸缩回
         Z04ExtPos : Bool := FALSE;   // 右防尘盖夹紧缸伸出
         Z04RetPos : Bool := TRUE;   // 右防尘盖夹紧缸缩回
         Z05Ext : Bool := FALSE;   // 供电抢打开
         Z05Ret : Bool := FALSE;   // 供电抢关闭
         Z06ExtPos : Bool := FALSE;   // 水泥板吹气打开
         Z06RetPos : Bool := TRUE;   // 水泥板吹气关闭
         Z07ExtPos : Bool := FALSE;   // 快换盘锁紧
         Z07RetPos : Bool := TRUE;   // 快换盘解锁
         CheckBit : Bool := FALSE;
         ClearHoleNum : Bool;   // 清零完成
         RobotBusy : Bool := FALSE;   // 机器人运行
         RobotReady : Bool := FALSE;   // 机器人启动
         RobotHome : Bool := FALSE;   // 机器人回原点
         RobotStop : Bool := FALSE;   // 机器人停止
         RobotClean : Bool := FALSE;   // 机器人清洁手动
         RobotTool : Bool := FALSE;   // 机器人换夹具手动
         RobotCheck : Bool := FALSE;   // 机器人校验手动
         RobotDrill : Bool := FALSE;   // 机器人钻孔手动
         Spare50 : Bool;
         Spare51 : Bool;
         Spare52 : Bool;
         Spare53 : Bool;
         ReqHeatMachine : Bool;   // 请求热机
         ToolPowerOn : Bool;
         Spare56 : Bool;
         Spare57 : Bool;
         RobotProgNo : Int := 16#00;   // 机器人反馈程序号
         PromptValue : Int;   // PromptValue
         HoleNo : Int := 0;   // 备用
         PowerCode : Int;   // 当前电源编码
         PosNo : Int;   // 当前打孔点位
         IoCode : Int;   // 当前信号编码
         ScrLen : Real;   // 当前钻孔深度
         CurrentPressure : Real;   // 当前压力
         Horizontal_OffSetY : Real;   // 当前水平Y工作坐标
         Horizontal_OffSetZ : Real;   // 当前水平Z工作坐标
         Download_OffSetY : Real;   // 当前垂直下Y工作坐标
         Download_OffSetX : Real;   // 当前垂直下X工作坐标
         Upload_OffSetY : Real;   // 当前垂直上Y工作坐标
         Upload_OffSetX : Real;   // 当前垂直上X工作坐标
         ScrTestLen : Real;   // 批头校验长度
         Layer : Int;   // 凿击层数
         Beer_info : Int;   // 错误信息
         Spare : Array[0..21] of Byte;
      END_STRUCT;
      Recv : Struct
         Heart : Bool := 0;   // 心跳
         EmmMode : Bool := 0;   // 紧急停止
         PcReady : Bool := 0;   // 上位机就绪
         PowerOff : Bool := 0;   // 枪关闭
         DataWriteDone : Bool;   // 参数写入完成
         ClearHoleNoReq : Bool;   // 请求清零孔数
         Spare4 : Bool;
         Spare5 : Bool;
         ParaWriteDone : Bool;   // 参数写入完成
         DrillStart : Bool;   // 进行打孔作业
         ChangeTool : Bool;   // 更换电锤
         WorkDone : Bool;   // 作业完成
         WorkStart : Bool;   // 作业开始
         HorizontalConfirm : Bool;   // 水平输入确认
         DownloadConfirm : Bool;   // 向下输入确认
         UploadConfirm : Bool;   // 向上输入确认
         Z01ExtTPPB : Bool := FALSE;   // 推力气缸伸出
         Z01RetTPPB : Bool := FALSE;   // 推力气缸缩回
         Z02ExtTPPB : Bool := FALSE;   // 辅助气缸伸出
         Z02RetTPPB : Bool := FALSE;   // 辅助气缸缩回
         Z03ExtTPPB : Bool := FALSE;   // 左防尘盖夹紧缸伸出
         Z03RetTPPB : Bool := FALSE;   // 左防尘盖夹紧缸缩回
         Z04ExtTPPB : Bool := FALSE;   // 右防尘盖夹紧缸伸出
         Z04RetTPPB : Bool := FALSE;   // 右防尘盖夹紧缸缩回
         Z05ExtTPPB : Bool := FALSE;   // 供电抢打开
         Z05RetTPPB : Bool := FALSE;   // 供电抢关闭
         Z06ExtTPPB : Bool := FALSE;   // 水泥板吹气打开
         Z06RetTPPB : Bool := FALSE;   // 水泥板吹气关闭
         Z07ExtTPPB : Bool := FALSE;   // 快换盘锁紧
         Z07RetTPPB : Bool := FALSE;   // 快换盘解锁
         Z01VentValveTPPB : Bool;   // 推力气缸中泄
         Z02VentValveTPPB : Bool;   // 辅助气缸中泄
         RobotStart : Bool := FALSE;   // 机器人启动
         RobotHoming : Bool := FALSE;   // 机器人回原点
         RobotStopTPPB : Bool := FALSE;   // 机器人停止
         CleanToolTPPB : Bool := FALSE;   // 机器人清洁手动
         ChangeToolTPPB : Bool := FALSE;   // 机器人换夹具手动
         CheckAiguilleTPPB : Bool := FALSE;   // 机器人校验手动
         RobotDrillTPPB : Bool := FALSE;   // 机器人钻孔手动
         Spare13 : Bool;
         ChangeHorizontalSlabDone : Bool := FALSE;   // 水平水泥板更换完成
         ChangeUploadSlabDone : Bool := FALSE;   // 垂直向上水泥板更换完成
         ChangeDownloadSlabDone : Bool := FALSE;   // 垂直向下水泥板更换完成
         PosNoClear : Bool;   // 打孔位清零
         ResHeatMachin : Bool;   // 热机完成
         Spare55 : Bool := 16#00;
         RobotPrigNo : Byte := 16#00;   // 输入程序号
         ChooseProgNo : Int := 0;   // 选择动作1水平2向下3向上4批头5力
         RunningNo : Int := 0;   // 流程数量
         Horizontal_OffSetY : Real := 0.0;   // 水平Y偏移量
         Horizontal_OffSetZ : Real;   // 水平Z偏移量
         Download_OffSetY : Real := 0.0;   // 向下Y偏移量
         Download_OffSetX : Real;   // 向下X偏移量
         Upload_OffSetY : Real := 0.0;   // 向上Y偏移量
         Current_1 : Real;   // 电流实时值1
         Current_2 : Real;   // 电流实时值2
         Layer : Int;   // 凿击层数
         DownSlabHeight : Int := 400;   // 向下水泥块厚度
         Voltage : Real;   // 电压
         Spare : Byte;
      END_STRUCT;
      Para : Struct
         DC_AC : Bool := 0;   // 交直流
         DrillDirection1 : Bool;   // 水平钻孔方向
         DrillDirection2 : Bool;   // 垂直向上钻孔方向
         DrillDirection3 : Bool;   // 垂直向下钻孔方向
         ProduceMode1 : Bool;   // 单钻
         ProduceMode2 : Bool;   // 锤钻
         ProduceMode3 : Bool;   // 单凿
         ControlMode : Bool;   // 自动结束方式：0-时间控制，1-孔数控制
         SwingOn : Bool;   // 摆动开
         DrillEndMode : Bool;   // 单个孔位结束模式：0-深度到达结束，1-时间到达结束
         DiamondVibCylinder : Bool;   // 水钻敲击功能启用
         spare_3 : Bool;
         spare_4 : Bool;
         spare_5 : Bool;
         spare_6 : Bool;
         spare_7 : Bool;
         IOFixtureNo : Byte := 16#00;   // 信号夹具号
         PowerFixtureNo : Byte;   // 电源夹具号
         TypeNo : Int := 0;   // 品种号
         WorkingFrequency : Int := 0;   // 单位Hz
         RobotSpeed : Int;   // 机器人运行速度
         DrillWidth : Real := 40.0;   // 钻孔宽度Y mm
         DrillDepth : Real := 90.0;   // 钻孔深度 mm
         HoleNum : Int;   // 钻孔数量
         Classification : Int := 0;   // 工作对象：1-水泥2-红砖-3轻质砖
         RestHours : DInt := 0;   // 单位S
         InputVoltage : Real := 0.0;   // 上位机使用，可以不发送
         InitialForce : Real := 0.0;   // 初始力 单位N
         ScrLen : Real := 120.0;   // 批头长度
         ZeroPos : Real := 1011.0;   // 枪校验原点坐标
         HorConcreteY : Real := 1200.0;   // 水平水泥板长
         HorConcreteZ : Real := 750.0;   // 水平水泥板宽
         UpConcreteY : Real := 1000.0;   // 垂直向上水泥板长
         UpConcreteX : Real := 700.0;   // 垂直向上水泥板宽
         DownConcreteY : Real := 1200.0;   // 垂直向下水泥板长
         DownConcreteX : Real := 800.0;   // 垂直向下水泥板宽
         ToolType : Int;   // 工具种类
         ToolModel : Int;   // 工具型号
         Angle : Real;   // 凿击角度
         SwingSpeed : Int;   // 摆动速度
         TimeOut : DInt;   // 单个打孔（凿击、锤、钻）作业的超时时间
         DrillTime : DInt;   // 凿击以时间为结束判断时有效
         CurrentMaxLimit : Real;   // 凿击电流上限
         CurrentMinLimit : Real;   // 凿击电流下限
         CurrentMinLimitTimeOut : DInt;   // 电流下限超时时间
         Auto_Force : Array[1..200] of Real;   // 曲线力
      END_STRUCT;
   END_VAR
BEGIN
   Send.Spare[0] := 16#00;
   Send.Spare[1] := 16#00;
   Send.Spare[2] := 16#00;
   Send.Spare[3] := 16#00;
   Send.Spare[4] := 16#00;
   Send.Spare[5] := 16#00;
   Send.Spare[6] := 16#00;
   Send.Spare[7] := 16#00;
   Send.Spare[8] := 16#00;
   Send.Spare[9] := 16#00;
   Send.Spare[10] := 16#00;
   Send.Spare[11] := 16#00;
END_DATA_BLOCK

// folder: 005_Component/Cooling Fan

DATA_BLOCK "DB2008_CoolingFan[DB2008]"   // DB13
{ S7_Optimized_Access := 'TRUE' }
VERSION : 0.1
// stored: InstanceOfName FB2008_CoolingFan
"FB2008_CoolingFan"
BEGIN
END_DATA_BLOCK

// folder: 006_ Visual Chiseling

DATA_BLOCK "DB2100 Modbus Value"   // DB2100
{ S7_Optimized_Access := 'FALSE' }
VERSION : 0.1
   VAR
      "PLC Para" : Struct
         "Status Word" : Word;   // PLC状态字
         "Time Word 1" : Word;   // PLC 年月日
         "Time Word 2" : Word;   // PLC分秒
         "Time Word 3" : Word;   // PLC时
         "Reserved Word 4" : Word;
         "Reserved Word 5" : Word;
         "Reserved Word 6" : Word;
         "Reserved Word 7" : Word;
         "Reserved Word 8" : Word;
         "Reserved Word 9" : Word;
         "Reserved Word 10" : Word;
         "Reserved Word 11" : Word;
         "Reserved Word 12" : Word;
         "Reserved Word 13" : Word;
         "Reserved Word 14" : Word;
         "Reserved Word 15" : Word;
         "Reserved Word 16" : Word;
         "Reserved Word 17" : Word;
         "Reserved Word 18" : Word;
         "Reserved Word 19" : Word;
         "Reserved Word 20" : Word;
         "Reserved Word 21" : Word;
         "Reserved Word 22" : Word;
         "Reserved Word 23" : Word;
         "Reserved Word 24" : Word;
         "Reserved Word 25" : Word;
         "Reserved Word 26" : Word;
         "Reserved Word 27" : Word;
         "Reserved Word 28" : Word;
         "Reserved Word 29" : Word;
         "Reserved Word 30" : Word;
         "Reserved Word 31" : Word;
      END_STRUCT;
      "ROS Para" : Struct
         "Status Word" : Word;   // ROS状态字
         "Time Word_1" : Word;   // ROS年月日
         "Time Word_2" : Word;   // ROS分秒
         "Time Word_3" : Word;   // ROS时
         "Sequence Word" : Word;   // 序列
         "PointNum Word" : Word;   // 坐标点数
         "PointPage Word" : Word;   // 坐标页码
         PointX_0 : Word;
         PointY_0 : Word;
         PointZ_0 : Word;
         PointA_0 : Word;
         PointB_0 : Word;
         PointC_0 : Word;
         PointX_1 : Word;
         PointY_1 : Word;
         PointZ_1 : Word;
         PointA_1 : Word;
         PointB_1 : Word;
         PointC_1 : Word;
         PointX_2 : Word;
         PointY_2 : Word;
         PointZ_2 : Word;
         PointA_2 : Word;
         PointB_2 : Word;
         PointC_2 : Word;
         PointX_3 : Word;
         PointY_3 : Word;
         PointZ_3 : Word;
         PointA_3 : Word;
         PointB_3 : Word;
         PointC_3 : Word;
         PointX_4 : Word;
         PointY_4 : Word;
         PointZ_4 : Word;
         PointA_4 : Word;
         PointB_4 : Word;
         PointC_4 : Word;
         PointX_5 : Word;
         PointY_5 : Word;
         PointZ_5 : Word;
         PointA_5 : Word;
         PointB_5 : Word;
         PointC_5 : Word;
         PointX_6 : Word;
         PointY_6 : Word;
         PointZ_6 : Word;
         PointA_6 : Word;
         PointB_6 : Word;
         PointC_6 : Word;
         PointX_7 : Word;
         PointY_7 : Word;
         PointZ_7 : Word;
         PointA_7 : Word;
         PointB_7 : Word;
         PointC_7 : Word;
         PointX_8 : Word;
         PointY_8 : Word;
         PointZ_8 : Word;
         PointA_8 : Word;
         PointB_8 : Word;
         PointC_8 : Word;
         PointX_9 : Word;
         PointY_9 : Word;
         PointZ_9 : Word;
         PointA_9 : Word;
         PointB_9 : Word;
         PointC_9 : Word;
         PointX_10 : Word;
         PointY_10 : Word;
         PointZ_10 : Word;
         PointA_10 : Word;
         PointB_10 : Word;
         PointC_10 : Word;
         PointX_11 : Word;
         PointY_11 : Word;
         PointZ_11 : Word;
         PointA_11 : Word;
         PointB_11 : Word;
         PointC_11 : Word;
         "Reserved Word_111" : Word;
         "Reserved Word_112" : Word;
         "Reserved Word_113" : Word;
         "Reserved Word_114" : Word;
         "Reserved Word_115" : Word;
         "Reserved Word_116" : Word;
         "Reserved Word_117" : Word;
         "Reserved Word_118" : Word;
         "Reserved Word_119" : Word;
         "Reserved Word_120" : Word;
         "Reserved Word_121" : Word;
         "Reserved Word_122" : Word;
         "Reserved Word_123" : Word;
         "Reserved Word_124" : Word;
         "Reserved Word_125" : Word;
         "Reserved Word_126" : Word;
      END_STRUCT;
   END_VAR
BEGIN
END_DATA_BLOCK

DATA_BLOCK "DB2300 Point Value"   // DB2300
{ S7_Optimized_Access := 'FALSE' }
VERSION : 0.1
   VAR
      Point : Array[0..23] of Struct
         X : Word;
         Y : Word;
         Z : Word;
         "A" : Word;
         "B" : Word;
         C : Word;
      END_STRUCT;
   END_VAR
BEGIN
END_DATA_BLOCK

DATA_BLOCK "DB2400 Visual Calibration"   // DB2400
{ S7_Optimized_Access := 'TRUE' }
VERSION : 0.1
   VAR
      VCALI_MODE : Bool;
      VCALI_STEP : Int;
   END_VAR
BEGIN
END_DATA_BLOCK

DATA_BLOCK "DB2500 Visual Chiseling"   // DB2500
{ S7_Optimized_Access := 'FALSE' }
VERSION : 0.1
   VAR
      "PLC Time" : DTL;
      "ROS Time" : DTL;
      PointNumtoRobot : Int;
      PointAddressOffset : Int;
      RosErrorNum : Int;
      VisualChiselRound : Int;
      VisualChiselingMode : Bool;
      VisualChiselingManual : Bool;
      VisualCameraStart : Bool;
      VisualCameraEnd : Bool;
      VisualChiselingStart : Bool;
      VisualChiselingEnd : Bool;
      ManualOpenCamCover : Bool;
      ManualCloseCamCover : Bool;
      ManualActivateCam : Bool;
      ManualRequestPhoto : Bool;
      AutoActivateCam : Bool;
      ROSCalculationFault : Bool;
      RosComFault : Bool;
      Page1_ConfirmInf : Bool;
      Page2_ConfirmInf : Bool;
      RobotRetHomeCmd_AllMode : Bool;
      Pulse : Array[0..31] of Bool;
      OffSet : Struct
         X : Word;
         Y : Word;
         Z : Word;
         "A" : Word;
         "B" : Word;
         C : Word;
      END_STRUCT;
      OffSetValue : Struct
         X : Real;
         Y : Real;
         Z : Real;
         "A" : Real;
         "B" : Real;
         C : Real;
      END_STRUCT;
      OffsetB_Radian : Real;
      OffsetB_SinB : Real;
      OffsetB_GravityComp : Real;
      VChiselCamRound : Int := -1;
      CalCamRound_Mid : Int;
      RestartModbus1 : Bool;
      RestartModbus2 : Bool;
      RestartModbus3 : Bool;
      RestartModbus4 : Bool;
      VChiselEndPos : Bool;
      VChiselComLock : Bool;   // 视觉通信流程锁，防止与力控通信冲突
      RCV_POINT_NUM : Word;
      VChiselCamLock : Bool;
   END_VAR
BEGIN
END_DATA_BLOCK

DATA_BLOCK "DB2600 FT Control"   // DB2600
{ S7_Optimized_Access := 'FALSE' }
VERSION : 0.1
   VAR
      FTControlMode : Bool;
      FTSensorRunning : Bool;
      FTControlRunning : Bool;
      FTControlBreak : Bool;   // quit when ft too large to protect system
      FTComLock : Bool;   // lock modbus when ft com.
      FTComError : Bool;
      FTStep : Int;   // 状态机
      FTActionCnt : Int;   // 调整次数
      Pulse : Array[0..7] of Bool;
      TarPoint_in : Array[0..0] of Struct
         X : Word;
         Y : Word;
         Z : Word;
         "A" : Word;
         "B" : Word;
         C : Word;
      END_STRUCT;
      TarPoint_out : Struct
         X : Real;
         Y : Real;
         Z : Real;
         "A" : Real;
         "B" : Real;
         C : Real;
      END_STRUCT;
   END_VAR
BEGIN
   // Pulse[0] : trigger ft sensor launch
   // Pulse[1] : trigger ft calibration
   // Pulse[2] : trigger ft control
   // Pulse[3] : trigger ft control action
   // Pulse[4] : trigger ft control quit
   // Pulse[5] : trigger ft sensor shutdown
   // Pulse[6] : trigger ft reset
END_DATA_BLOCK

DATA_BLOCK "DB2700 Visual Point Reset"   // DB2700
{ S7_Optimized_Access := 'FALSE' }
VERSION : 0.1
   VAR
      "Modbus Value" : Struct
         PointX_0 : Word;
         PointY_0 : Word;
         PointZ_0 : Word;
         PointA_0 : Word;
         PointB_0 : Word;
         PointC_0 : Word;
         PointX_1 : Word;
         PointY_1 : Word;
         PointZ_1 : Word;
         PointA_1 : Word;
         PointB_1 : Word;
         PointC_1 : Word;
         PointX_2 : Word;
         PointY_2 : Word;
         PointZ_2 : Word;
         PointA_2 : Word;
         PointB_2 : Word;
         PointC_2 : Word;
         PointX_3 : Word;
         PointY_3 : Word;
         PointZ_3 : Word;
         PointA_3 : Word;
         PointB_3 : Word;
         PointC_3 : Word;
         PointX_4 : Word;
         PointY_4 : Word;
         PointZ_4 : Word;
         PointA_4 : Word;
         PointB_4 : Word;
         PointC_4 : Word;
         PointX_5 : Word;
         PointY_5 : Word;
         PointZ_5 : Word;
         PointA_5 : Word;
         PointB_5 : Word;
         PointC_5 : Word;
         PointX_6 : Word;
         PointY_6 : Word;
         PointZ_6 : Word;
         PointA_6 : Word;
         PointB_6 : Word;
         PointC_6 : Word;
         PointX_7 : Word;
         PointY_7 : Word;
         PointZ_7 : Word;
         PointA_7 : Word;
         PointB_7 : Word;
         PointC_7 : Word;
         PointX_8 : Word;
         PointY_8 : Word;
         PointZ_8 : Word;
         PointA_8 : Word;
         PointB_8 : Word;
         PointC_8 : Word;
         PointX_9 : Word;
         PointY_9 : Word;
         PointZ_9 : Word;
         PointA_9 : Word;
         PointB_9 : Word;
         PointC_9 : Word;
         PointX_10 : Word;
         PointY_10 : Word;
         PointZ_10 : Word;
         PointA_10 : Word;
         PointB_10 : Word;
         PointC_10 : Word;
         PointX_11 : Word;
         PointY_11 : Word;
         PointZ_11 : Word;
         PointA_11 : Word;
         PointB_11 : Word;
         PointC_11 : Word;
         PointX_12 : Word;
         PointY_12 : Word;
         PointZ_12 : Word;
         PointA_12 : Word;
         PointB_12 : Word;
         PointC_12 : Word;
         PointX_13 : Word;
         PointY_13 : Word;
         PointZ_13 : Word;
         PointA_13 : Word;
         PointB_13 : Word;
         PointC_13 : Word;
         PointX_14 : Word;
         PointY_14 : Word;
         PointZ_14 : Word;
         PointA_14 : Word;
         PointB_14 : Word;
         PointC_14 : Word;
         PointX_15 : Word;
         PointY_15 : Word;
         PointZ_15 : Word;
         PointA_15 : Word;
         PointB_15 : Word;
         PointC_15 : Word;
         PointX_16 : Word;
         PointY_16 : Word;
         PointZ_16 : Word;
         PointA_16 : Word;
         PointB_16 : Word;
         PointC_16 : Word;
         PointX_17 : Word;
         PointY_17 : Word;
         PointZ_17 : Word;
         PointA_17 : Word;
         PointB_17 : Word;
         PointC_17 : Word;
         PointX_18 : Word;
         PointY_18 : Word;
         PointZ_18 : Word;
         PointA_18 : Word;
         PointB_18 : Word;
         PointC_18 : Word;
         PointX_19 : Word;
         PointY_19 : Word;
         PointZ_19 : Word;
         PointA_19 : Word;
         PointB_19 : Word;
         PointC_19 : Word;
         PointX_20 : Word;
         PointY_20 : Word;
         PointZ_20 : Word;
         PointA_20 : Word;
         PointB_20 : Word;
         PointC_20 : Word;
         PointX_21 : Word;
         PointY_21 : Word;
         PointZ_21 : Word;
         PointA_21 : Word;
         PointB_21 : Word;
         PointC_21 : Word;
         PointX_22 : Word;
         PointY_22 : Word;
         PointZ_22 : Word;
         PointA_22 : Word;
         PointB_22 : Word;
         PointC_22 : Word;
         PointX_23 : Word;
         PointY_23 : Word;
         PointZ_23 : Word;
         PointA_23 : Word;
         PointB_23 : Word;
         PointC_23 : Word;
      END_STRUCT;
   END_VAR
BEGIN
END_DATA_BLOCK

// folder: System blocks/Program resources

DATA_BLOCK "Timer_Modbus1"   // DB2
{ S7_Optimized_Access := 'TRUE' }
AUTHOR : Simatic
FAMILY : IEC
NAME : IEC_TMR
VERSION : 1.0
// stored: InstanceOfName IEC_TIMER
"IEC_TIMER"
BEGIN
END_DATA_BLOCK

DATA_BLOCK "Timer_Modbus2"   // DB3
{ S7_Optimized_Access := 'TRUE' }
AUTHOR : Simatic
FAMILY : IEC
NAME : IEC_TMR
VERSION : 1.0
// stored: InstanceOfName IEC_TIMER
"IEC_TIMER"
BEGIN
END_DATA_BLOCK

DATA_BLOCK "Timer_Modbus3"   // DB4
{ S7_Optimized_Access := 'TRUE' }
AUTHOR : Simatic
FAMILY : IEC
NAME : IEC_TMR
VERSION : 1.0
// stored: InstanceOfName IEC_TIMER
"IEC_TIMER"
BEGIN
END_DATA_BLOCK

DATA_BLOCK "Timer_ParaWriteOuttime"   // DB5
{ S7_Optimized_Access := 'TRUE' }
AUTHOR : Simatic
FAMILY : IEC
NAME : IEC_TMR
VERSION : 1.0
// stored: InstanceOfName IEC_TIMER
"IEC_TIMER"
BEGIN
END_DATA_BLOCK

DATA_BLOCK "Timer_DownChiselEnd"   // DB6
{ S7_Optimized_Access := 'TRUE' }
AUTHOR : Simatic
FAMILY : IEC
NAME : IEC_TMR
VERSION : 1.0
// stored: InstanceOfName IEC_TIMER
"IEC_TIMER"
BEGIN
END_DATA_BLOCK

DATA_BLOCK "Timer_RecvEmmMode"   // DB8
{ S7_Optimized_Access := 'TRUE' }
AUTHOR : Simatic
FAMILY : IEC
NAME : IEC_TMR
VERSION : 1.0
// stored: InstanceOfName IEC_TIMER
"IEC_TIMER"
BEGIN
END_DATA_BLOCK

DATA_BLOCK "Timer_ft_bringup"   // DB9
{ S7_Optimized_Access := 'TRUE' }
AUTHOR : Simatic
FAMILY : IEC
NAME : IEC_TMR
VERSION : 1.0
// stored: InstanceOfName IEC_TIMER
"IEC_TIMER"
BEGIN
END_DATA_BLOCK

DATA_BLOCK "Timer_ft_calib"   // DB10
{ S7_Optimized_Access := 'TRUE' }
AUTHOR : Simatic
FAMILY : IEC
NAME : IEC_TMR
VERSION : 1.0
// stored: InstanceOfName IEC_TIMER
"IEC_TIMER"
BEGIN
END_DATA_BLOCK

DATA_BLOCK "Timer_ft_ctrl"   // DB11
{ S7_Optimized_Access := 'TRUE' }
AUTHOR : Simatic
FAMILY : IEC
NAME : IEC_TMR
VERSION : 1.0
// stored: InstanceOfName IEC_TIMER
"IEC_TIMER"
BEGIN
END_DATA_BLOCK

DATA_BLOCK "Timer_CamCalc"   // DB12
{ S7_Optimized_Access := 'TRUE' }
AUTHOR : Simatic
FAMILY : IEC
NAME : IEC_TMR
VERSION : 1.0
// stored: InstanceOfName IEC_TIMER
"IEC_TIMER"
BEGIN
END_DATA_BLOCK

DATA_BLOCK "Timer05_ChiselStart"   // DB2505
{ S7_Optimized_Access := 'TRUE' }
AUTHOR : Simatic
FAMILY : IEC
NAME : IEC_TMR
VERSION : 1.0
// stored: InstanceOfName IEC_TIMER
"IEC_TIMER"
BEGIN
END_DATA_BLOCK

DATA_BLOCK "Timer10_ChiselCam"   // DB2510
{ S7_Optimized_Access := 'TRUE' }
AUTHOR : Simatic
FAMILY : IEC
NAME : IEC_TMR
VERSION : 1.0
// stored: InstanceOfName IEC_TIMER
"IEC_TIMER"
BEGIN
END_DATA_BLOCK

DATA_BLOCK "Timer15_ChiselCom"   // DB2515
{ S7_Optimized_Access := 'TRUE' }
AUTHOR : Simatic
FAMILY : IEC
NAME : IEC_TMR
VERSION : 1.0
// stored: InstanceOfName IEC_TIMER
"IEC_TIMER"
BEGIN
END_DATA_BLOCK

DATA_BLOCK "Timer20_ChiselPage1"   // DB2520
{ S7_Optimized_Access := 'TRUE' }
AUTHOR : Simatic
FAMILY : IEC
NAME : IEC_TMR
VERSION : 1.0
// stored: InstanceOfName IEC_TIMER
"IEC_TIMER"
BEGIN
END_DATA_BLOCK

DATA_BLOCK "Timer25_ChiselPage2"   // DB2525
{ S7_Optimized_Access := 'TRUE' }
AUTHOR : Simatic
FAMILY : IEC
NAME : IEC_TMR
VERSION : 1.0
// stored: InstanceOfName IEC_TIMER
"IEC_TIMER"
BEGIN
END_DATA_BLOCK

DATA_BLOCK "Timer30_ChiselStepEnd"   // DB2530
{ S7_Optimized_Access := 'TRUE' }
AUTHOR : Simatic
FAMILY : IEC
NAME : IEC_TMR
VERSION : 1.0
// stored: InstanceOfName IEC_TIMER
"IEC_TIMER"
BEGIN
END_DATA_BLOCK

DATA_BLOCK "Timer35_ChiselEnd"   // DB2535
{ S7_Optimized_Access := 'TRUE' }
AUTHOR : Simatic
FAMILY : IEC
NAME : IEC_TMR
VERSION : 1.0
// stored: InstanceOfName IEC_TIMER
"IEC_TIMER"
BEGIN
END_DATA_BLOCK

DATA_BLOCK "Timer_CylinderBack_Hor"   // DB3000
{ S7_Optimized_Access := 'TRUE' }
AUTHOR : Simatic
FAMILY : IEC
NAME : IEC_TMR
VERSION : 1.0
// stored: InstanceOfName IEC_TIMER
"IEC_TIMER"
BEGIN
END_DATA_BLOCK

DATA_BLOCK "Timer_RobotPry_Hor"   // DB3010
{ S7_Optimized_Access := 'TRUE' }
AUTHOR : Simatic
FAMILY : IEC
NAME : IEC_TMR
VERSION : 1.0
// stored: InstanceOfName IEC_TIMER
"IEC_TIMER"
BEGIN
END_DATA_BLOCK

DATA_BLOCK "Timer_CylinderBack_Down"   // DB3020
{ S7_Optimized_Access := 'TRUE' }
AUTHOR : Simatic
FAMILY : IEC
NAME : IEC_TMR
VERSION : 1.0
// stored: InstanceOfName IEC_TIMER
"IEC_TIMER"
BEGIN
END_DATA_BLOCK

DATA_BLOCK "Timer_RobotPry_Down"   // DB3030
{ S7_Optimized_Access := 'TRUE' }
AUTHOR : Simatic
FAMILY : IEC
NAME : IEC_TMR
VERSION : 1.0
// stored: InstanceOfName IEC_TIMER
"IEC_TIMER"
BEGIN
END_DATA_BLOCK

DATA_BLOCK "Counter_VChiselRound"   // DB3040
{ S7_Optimized_Access := 'TRUE' }
AUTHOR : Simatic
FAMILY : IEC
NAME : CNTR
VERSION : 1.0
// stored: InstanceOfName IEC_COUNTER
"IEC_COUNTER"
BEGIN
END_DATA_BLOCK

DATA_BLOCK "Timer_DrilEndPos"   // DB3050
{ S7_Optimized_Access := 'TRUE' }
AUTHOR : Simatic
FAMILY : IEC
NAME : IEC_TMR
VERSION : 1.0
// stored: InstanceOfName IEC_TIMER
"IEC_TIMER"
BEGIN
END_DATA_BLOCK

DATA_BLOCK "Timer_ChangeChiselArea"   // DB3060
{ S7_Optimized_Access := 'TRUE' }
AUTHOR : Simatic
FAMILY : IEC
NAME : IEC_TMR
VERSION : 1.0
// stored: InstanceOfName IEC_TIMER
"IEC_TIMER"
BEGIN
END_DATA_BLOCK

// folder: (top level)

FUNCTION_BLOCK "FB1001_SysMode"   // FB1001, SCL
{ S7_Optimized_Access := 'TRUE' }
// ============================================================
//  Block: FB1001_SysMode
//  ============================================================
//  编号：FB1001
//  原始语言：LAD（规则翻译为 SCL）
//  含义：***********************************************************************************************************************************************************************************不能更改************************************************************************************************************************************************************
   VAR_INPUT
      I_OkToStartNew : Bool;   // 输入参数
      iEMOK : Bool;   // 输入参数
      iAirPressOK : Bool;   // 输入参数
      iManMode : Bool;   // 输入参数
      iAutoMode : Bool;   // 输入参数
      iAutoModeStart : Bool;   // 输入参数
      iBeeperQuiet : Bool;   // 输入参数
      iErrRst : Bool;   // 输入参数
      iStartL : Bool;   // 输入参数
      iStartR : Bool;   // 输入参数
      I_ErrPresent : Bool;   // 输入参数
      I_ErrAutoReset : Bool;   // 输入参数
      I_AutoRuning : Bool;   // 输入参数
      I_HomeIng : Bool;   // 输入参数
      I_AllStationInHomePos : Bool;   // 输入参数
      iHomeMode : Bool;   // 输入参数
      I_SP2 : Bool;   // 输入参数
   END_VAR
   VAR_OUTPUT
      oTLBlue : Bool;   // 输出参数
      oTLYel : Bool;   // 输出参数
      oTLGreen : Bool;   // 输出参数
      oTLRed : Bool;   // 输出参数
      oTLWhite : Bool;   // 输出参数
      oPanelG : Bool;   // 输出参数
      oPanelRed : Bool;   // 输出参数
      oBeeper : Bool;   // 输出参数
      oLightingLampClose : Bool;   // 输出参数
      oEMErr : Bool;   // 输出参数
      oPressErr : Bool;   // 输出参数
      oErrToBeRst : Bool;   // 输出参数
      oStartAutoModePrompt : Bool;   // 输出参数
      oAutoModeOffPrompt : Bool;   // 输出参数
      oEmptyMode : Bool;   // 输出参数
      oStepMode : Bool;   // 输出参数
      oModeFromTP : Bool;   // 输出参数
   END_VAR
   VAR
      TP_Cmd : Word;   // 静态变量
      Cmd : Struct   // 静态变量
         ClearCounter : Bool;   // 静态变量
         SetTime : Bool;   // 静态变量
      END_STRUCT;
      At_Cmd : Word;   // 静态变量
      Cylinder_Index : Int := 1;   // 从1开始
      SysMode_Station_Index : Int := 1;   // 静态变量
      Sys_Time : Struct   // 静态变量
         CurPLCTime : DTL := DTL#2015-03-21-17:23:15;   // 静态变量
         SetPLCTimeTP : DTL;   // 静态变量
      END_STRUCT;
      SubSysMode : "FB1002_subSysMode";   // 静态变量
      OUT : Struct   // 静态变量
         LampTest : Bool;   // 静态变量
         oPanelHome : Bool;   // 静态变量
         sp : Word;   // 静态变量
      END_STRUCT;
      Mode : Struct   // 静态变量
         ManMode : Bool;   // 静态变量
         MastMode : Bool;   // 静态变量
         StepMode : Bool;   // 静态变量
         AutoMode : Bool;   // 静态变量
         EMMode : Bool;   // 静态变量
         PressLowMode : Bool;   // 静态变量
         sp_1 : Bool;   // 静态变量
         sp_2 : Bool;   // 静态变量
         ASMode : Bool;   // 静态变量
         ASMMode : Bool;   // 静态变量
         AllMode : Bool;   // 静态变量
         HomeCmd : Bool;   // 静态变量
         ErrRst : Bool;   // 静态变量
         StartPls : Bool;   // 静态变量
         StepPls : Bool;   // 静态变量
         StartLeftPls : Bool;   // 静态变量
         StartRightPls : Bool;   // 静态变量
         StepLeftPls : Bool;   // 静态变量
         StepRightPls : Bool;   // 静态变量
         ManModePls : Bool;   // 静态变量
         AllModePls : Bool;   // 静态变量
         sp : DWord;   // 静态变量
      END_STRUCT;
      TPPB : Struct   // 静态变量
         EmptyMode : Bool;   // 静态变量
         Bypass : Bool;   // 静态变量
         STAT6 : Bool;   // 静态变量
         STAT5 : Bool;   // 静态变量
         STAT4 : Bool;   // 静态变量
         STAT3 : Bool;   // 静态变量
         STAT2 : Bool;   // 静态变量
         STAT1 : Bool;   // 静态变量
         LampTest : Bool;   // 静态变量
         Home : Bool;   // 静态变量
         StepMode : Bool;   // 静态变量
         ErrRst : Bool;   // 静态变量
         LampCtrol : Bool;   // 静态变量
         Quiet : Bool;   // 静态变量
         opModeFromTP : Bool;   // 静态变量
         sp : DWord;   // 静态变量
      END_STRUCT;
      Status : Struct   // 静态变量
         HomePos : Bool;   // 静态变量
         HomeIng : Bool;   // 静态变量
         AutoRunning : Bool;   // 静态变量
         ErrPresent : Bool;   // 静态变量
         AutoModeStarted : Bool;   // 静态变量
      END_STRUCT;
      TPSetPageNo : Int;   // 静态变量
      TPCurPageType : Int;   // 静态变量
      TPCurSubPage : Int;   // 静态变量
      IO_FromTP : Struct   // 静态变量
         spbyte : Byte;   // 静态变量
         EMOK : Bool;   // 静态变量
         AirPressOK : Bool;   // 静态变量
         ManMode : Bool;   // 静态变量
         AutoMode : Bool;   // 静态变量
         AutoModeStart : Bool;   // 静态变量
         ErrRst : Bool;   // 静态变量
         StartLeft : Bool;   // 静态变量
         StartRight : Bool;   // 静态变量
      END_STRUCT;
      IO_Cur : Struct   // 静态变量
         spbyte : Byte;   // 静态变量
         EMOK : Bool;   // 静态变量
         AirPressOK : Bool;   // 静态变量
         ManMode : Bool;   // 静态变量
         AutoMode : Bool;   // 静态变量
         AutoModeStart : Bool;   // 静态变量
         ErrRst : Bool;   // 静态变量
         StartLeft : Bool;   // 静态变量
         StartRight : Bool;   // 静态变量
      END_STRUCT;
      ModeDT : Struct   // 静态变量
         ManMode1 : Bool;   // 静态变量
         ManMode2 : Bool;   // 静态变量
         AutoMode1 : Bool;   // 静态变量
         AutoMode2 : Bool;   // 静态变量
         MastMode1 : Bool;   // 静态变量
         MastMode2 : Bool;   // 静态变量
         HomeCmd1 : Bool;   // 静态变量
         HomeCmd2 : Bool;   // 静态变量
         HomeCmd3 : Bool;   // 静态变量
         HomeCmd4 : Bool;   // 静态变量
         ErrLampOn01 : Bool;   // 静态变量
         ErrLampOn02 : Bool;   // 静态变量
      END_STRUCT;
      Aux : Struct   // 静态变量
         BeeperON_Keep : Bool;   // 静态变量
         BeeperOn : Bool;   // 静态变量
         BeeperOnPls : Bool;   // 静态变量
         ManMode : Bool;   // 静态变量
         ManModePls : Bool;   // 静态变量
         AutoMode : Bool;   // 静态变量
         AutoModePls : Bool;   // 静态变量
         ModeChangePlsHW : Bool;   // 静态变量
         AutoRunningPls : Bool;   // 静态变量
         OKPartPromptPls : Bool;   // 静态变量
         NGPartPromptPls : Bool;   // 静态变量
         ManModeOn : Bool;   // 静态变量
         AllModeOn : Bool;   // 静态变量
         AutoModeStartBtnPls : Bool;   // 静态变量
         AutoModeOnPls : Bool;   // 静态变量
         AutoModeOffCmd : Bool;   // 静态变量
         TPCurSubPage : Int;   // 静态变量
      END_STRUCT;
      Start1DT1 : IEC_TIMER;   // 静态变量
      Start1DT2 : IEC_TIMER;   // 静态变量
      Start2DT1 : IEC_TIMER;   // 静态变量
      Start2DT2 : IEC_TIMER;   // 静态变量
      xArray_SP : Array[0..91] of Byte;   // 静态变量
      lastByteAddr : Byte;   // 静态变量
      PT : Time;   // 静态变量
      ET : Time;   // 静态变量
      IN : Bool;   // 静态变量
      Q : Bool;   // 静态变量
   END_VAR
   VAR_TEMP
      RetVal : Int;   // 临时变量
      T_Bool : Bool;   // 临时变量
   END_VAR
BEGIN

   // ---------- 网络 1 ----------
   // 标题：PLC Time;
   // 含义：调用计数器实例 RD_SYS_T（上升沿计数，当前值写入 CV）
   #RetVal := RD_SYS_T(#Sys_Time.CurPLCTime);
   // 含义：调用定时器实例 WR_SYS_T
   IF #Cmd.SetTime THEN
       #RetVal := WR_SYS_T(#Sys_Time.SetPLCTimeTP);
   END_IF;

   // ---------- 网络 2 ----------
   // 标题：读取系统时间，为了做定时器
   // 注释：***********************************************************************************************************************************************************************************不能更改************************************************************************************************************************************************************
   // 含义：将 #Sys_Time.CurPLCTime; (* T_CONV DTL → Time_Of_Day *) 赋给 "SyS_Time"
   "SyS_Time" := DTL_TO_TOD(#Sys_Time.CurPLCTime);

   // ---------- 网络 3 ----------
   // 标题：初始化SysMode_Station_Index
   // 含义：条件 "DB1000_StdSignal".PLS.InitialPls 成立时，将 1 传送到 #Cylinder_Index
   IF "DB1000_StdSignal".PLS.InitialPls THEN
       #Cylinder_Index := 1;
   END_IF;
   // 含义：条件 "DB1000_StdSignal".PLS.InitialPls 成立时，将 1 传送到 #SysMode_Station_Index
   IF "DB1000_StdSignal".PLS.InitialPls THEN
       #SysMode_Station_Index := 1;
   END_IF;

   // ---------- 网络 4 ----------
   // 标题：转移触摸屏常用命令
   // 含义：将 #TP_Cmd 赋给 #At_Cmd
   #At_Cmd := #TP_Cmd;
   // 含义：将 0 赋给 #TP_Cmd
   #TP_Cmd := 0;

   // ---------- 网络 5 ----------
   // 标题：OPK020工位的模式
   // 含义：调用定时器实例 #SubSysMode
   #SubSysMode(iAirPressOK := "IAirPressOK",
               iManMode := "IMan",
               iAutoMode := "IAuto",
               iAutoModeStart := "IAutoModeStart",
               iErrRst := "IErrRst",
               I_ErrPresent := "DB1140_Message".o_Err,
               I_AutoRuning := "DB1060_AutoStep".Status.Running,
               I_HomeIng := "DB1040_HomePos".Status.Running,
               I_AllStationInHomePos := "DB1040_HomePos".Status.AllStationInHomePos,
               oTLBlue => "QTLB",
               oTLYel => "QTLY",
               oTLGreen => "QTLG",
               oTLRed => "QTLR",
               oTLWhite => "QTLW",
               oPanelG => "QPanelG",
               oPanelRed => "QPanelRed",
               oBeeper => "QBeeper",
               oLightingLampClose => "QLampCtr",
               oEMErr => "DB1148_PromptBeeper".Public.EMING,
               oPressErr => "DB1148_PromptBeeper".Public.AirPressureLow,
               oStartAutoModePrompt => "DB1146_PromptFree".Public.AutoModeNotStarted,
               oAutoModeOffPrompt => "DB1146_PromptFree".Public.AutoModeOffPrompt,
               oEmptyMode => "DB1146_PromptFree".Public.EmptyMode,
               oStepMode => "DB1146_PromptFree".Public.StepMode,
               oModeFromTP => "DB1146_PromptFree".Public.WaitPcCommond);

